// TwinCAT 3 PLC project PLCLibrary
// Title: LPLC
// Company: LPLC
// Author: Arya Farzin
// ProjectVersion: 2.2.0
// Description: LPLC - standardized TwinCAT 3 device, motion and machine function blocks (companion PLC library to lhmi). MIT License.
// ProgramVersion: 3.1.4026.17
// libraries:
//   Tc2_MC2, * (Beckhoff Automation GmbH)
//   Tc2_MC2_Camming, * (Beckhoff Automation GmbH)
//   Tc2_ModbusSrv, * (Beckhoff Automation GmbH)
//   Tc2_Standard, * (Beckhoff Automation GmbH)
//   Tc2_SUPS, * (Beckhoff Automation GmbH)
//   Tc2_System, * (Beckhoff Automation GmbH)
//   Tc2_Utilities, * (Beckhoff Automation GmbH)
//   Tc3_EventLogger, * (Beckhoff Automation GmbH)
//   Tc3_IotBase, * (Beckhoff Automation GmbH)
//   Tc3_JsonXml, * (Beckhoff Automation GmbH)
// project tree:
//   DUTs/Abstract/abs_fb_Device/ ST_Device_HMI_Interface.TcDUT
//   DUTs/Abstract/abs_fb_stateDevice/ ST_StateDevice_HMI_Commands.TcDUT, ST_StateDevice_HMI_Interface.TcDUT, ST_StateDevice_HMI_Status.TcDUT
//   DUTs/Abstract/abs_fb_MachineFlow/ ST_MachineFlow_HMI_Status.TcDUT, ST_MachineFlow_Step.TcDUT, ST_MachineFlow_Transition.TcDUT
//   DUTs/Devices/fb_Dev_StackLight3SegHV_BannerTL50Pro/ EN_Banner_TL503Pro_Animation.TcDUT, EN_Banner_TL503Pro_Colors.TcDUT, ST_Banner_TL503Pro.TcDUT, ST_Banner_TL503Pro_Raw.TcDUT
//   DUTs/Comm/fb_Modbus_Driver/ E_DriverState.TcDUT, E_MBArea.TcDUT, E_MBDataType.TcDUT, E_SignalQuality.TcDUT, E_WordOrder.TcDUT, ST_BitRegisterRmw.TcDUT, ST_MBDeviceStatus.TcDUT, ST_MBReadResult.TcDUT, ST_MBSignalConfig.TcDUT, ST_MBWriteData.TcDUT, ST_ParsedSignal.TcDUT, ST_ReadBlock.TcDUT, ST_WriteBlock.TcDUT
//   DUTs/Comm/fb_MQTT_Connector/ E_MQTT_Direction.TcDUT, E_MQTT_PublishMode.TcDUT, E_MQTT_SignalType.TcDUT, ST_MQTT_Signal.TcDUT
//   DUTs/Devices/fb_Dev_AnalogSensor/ ST_AnalogSensor_Diag.TcDUT, ST_AnalogSensor_HMI_Interface.TcDUT
//   DUTs/Devices/fb_Dev_IsolationMonitor/ ST_IsoMon_DeviceSignals.TcDUT, ST_IsoMon_HMI_Interface.TcDUT, ST_IsoMon_MBIF.TcDUT
//   DUTs/Devices/fb_Dev_PSU_ITECH/ ST_ITECH_DCMeter.TcDUT, ST_ITECH_DCSource.TcDUT, ST_ITECH_DeviceSignals.TcDUT, ST_ITECH_HMI_DeviceSignals.TcDUT, ST_ITECH_Protection.TcDUT, ST_ITECH_QuestionRegister.TcDUT, ST_ITECH_SetConfigs.TcDUT, ST_ITECH_SoftwareFaults.TcDUT, ST_ITECH_SystemStatus.TcDUT
//   DUTs/Devices/fb_Dev_Pump_ABBACS580/ ST_Pump_ABBACS580_HMI_Interface.TcDUT
//   DUTs/Devices/fb_Dev_Pump_SPAL/ EN_Pump_SPAL_Operating_Status.TcDUT, EN_Pump_SPAL_PumpError.TcDUT, EN_Pump_SPAL_ServiceIndicator.TcDUT, ST_Pump_SPAL_CAN_Inputs.TcDUT, ST_Pump_SPAL_CAN_Outputs.TcDUT, ST_Pump_SPAL_HMI_Interface.TcDUT
//   DUTs/Devices/fb_Dev_Actuator/ ST_Actuator_HMI_Interface.TcDUT
//   DUTs/Devices/fb_Dev_VFD_ABBACS580/ ST_VFD_ABBACS580_HMI_Interface.TcDUT, ST_VFD_ABBACS580_Telemetry.TcDUT
//   DUTs/Devices/fb_Dev_VFD_DuraPulse/ ST_VFD_DuraPulse_HMI_Interface.TcDUT, ST_VFD_DuraPulse_Telemetry.TcDUT
//   DUTs/fb_Axis/ E_Axis_BufferMode.TcDUT, E_Axis_JogSource.TcDUT, E_Axis_Mode.TcDUT, E_Axis_UnitType.TcDUT, ST_Axis_HMI_Commands.TcDUT, ST_Axis_HMI_Config.TcDUT, ST_Axis_HMI_Interface.TcDUT, ST_Axis_HMI_Status.TcDUT, ST_Axis_MoveDefinition.TcDUT
//   DUTs/Camming/fb_CamCoupler/ E_CamCoupler_State.TcDUT, ST_CamCoupler_HMI_Commands.TcDUT, ST_CamCoupler_HMI_Config.TcDUT, ST_CamCoupler_HMI_Interface.TcDUT, ST_CamCoupler_HMI_Status.TcDUT
//   DUTs/Camming/fb_CamTeach/ E_CamTeach_Interp.TcDUT, E_CamTeach_State.TcDUT, ST_CamTeach_HMI_Commands.TcDUT, ST_CamTeach_HMI_Config.TcDUT, ST_CamTeach_HMI_Interface.TcDUT, ST_CamTeach_HMI_Status.TcDUT, ST_CamTeach_Point.TcDUT
//   DUTs/Devices/fb_Dev_StripLight_BannerWLS15Pro/ E_BannerWLS15Pro_Animation.TcDUT, E_BannerWLS15Pro_Color.TcDUT, E_BannerWLS15Pro_Direction.TcDUT, E_BannerWLS15Pro_Intensity.TcDUT, E_BannerWLS15Pro_PulsePattern.TcDUT, E_BannerWLS15Pro_ScrollBounceStyle.TcDUT, E_BannerWLS15Pro_Speed.TcDUT, ST_Banner_WLS15PXRGB0220DSKQP_RunMode_Outputs.TcDUT
//   DUTs/Devices/fb_Dev_XPendant/ ST_XPendant_Axis.TcDUT, ST_XPendant_HMI_Interface.TcDUT, ST_XPendant_HMI_Status.TcDUT, ST_XPendant_In.TcDUT
//   DUTs/Common/ ST_Bits.TcDUT, U_ByteToLReal.TcDUT, U_UINT16.TcDUT, U_USINT.TcDUT
//   DUTs/Devices/fb_Dev_ControlValve_Modulating/ ST_ControlValve_Modulating_HMI_Interface.TcDUT
//   DUTs/fb_IO_EL6751_Bus_Status/ ST_EL6751_Bus_State.TcDUT, ST_EL6751_Bus_State_Parsed.TcDUT
//   DUTs/fb_Interlock/ ST_Interlock.TcDUT, ST_Interlock_HMI_Interface.TcDUT
//   DUTs/fb_Permissive/ ST_Permissive.TcDUT, ST_Permissive_HMI_Interface.TcDUT
//   DUTs/fb_Machine/ ST_Machine_HMI_Interface.TcDUT
//   DUTs/Comm/ ST_Modbus_Commands.TcDUT, ST_Modbus_Device_Config.TcDUT
//   POUs/FBs/Abstract/ abs_fb_Device.TcPOU, abs_fb_MachineFlow.TcPOU, abs_fb_stateDevice.TcPOU
//   POUs/FBs/Comm/ fb_Modbus_Driver.TcPOU, fb_MQTT_Connector.TcPOU
//   POUs/FBs/ fb_WriteDataToFile.TcPOU, fb_Axis.TcPOU, fb_FaultMonitor.TcPOU, fb_HmiEventLog.TcPOU, fb_Interlock.TcPOU, fb_Permissive.TcPOU, fb_IO_EL6751_Bus_Status.TcPOU, fb_Machine.TcPOU, fb_PID_Clamping.TcPOU, fb_RampGenerator.TcPOU, fb_SampleBuffer.TcPOU, fb_TimeAverage.TcPOU
//   POUs/FBs/Devices/ fb_Dev_Actuator.TcPOU, fb_Dev_XPendant.TcPOU, fb_Dev_AnalogSensor.TcPOU, fb_Dev_AnalogSensor_Accelerometer.TcPOU, fb_Dev_AnalogSensor_CurrentTransducer.TcPOU, fb_Dev_AnalogSensor_ELM_10x.TcPOU, fb_Dev_AnalogSensor_ELM_10x_CurrentTransducer.TcPOU, fb_Dev_ControlValve_Modulating_INT.TcPOU, fb_Dev_Pump_ABBACS580.TcPOU, fb_Dev_VFD_ABBACS580.TcPOU, fb_Dev_VFD_DuraPulse.TcPOU, fb_Dev_WebRelay.TcPOU, fb_Dev_ControlValve_Modulating.TcPOU, fb_Dev_ControlValve_Modulating_REAL.TcPOU, fb_Dev_IsolationMonitor.TcPOU, fb_Dev_Machine.TcPOU, fb_Dev_PSU_ITECH.TcPOU, fb_Dev_Pump_SPAL.TcPOU, fb_Dev_StackLight3SegHV_BannerTL50Pro.TcPOU, fb_Dev_StripLight_BannerWLS15Pro.TcPOU
//   POUs/FBs/Camming/ fb_CamCoupler.TcPOU, fb_CamTeach.TcPOU, fb_CamTeachFile.TcPOU
//   POUs/FC/ F_AddToArray_String.TcPOU, F_AnalogToEngUnit.TcPOU, F_RemoveFromArray_String.TcPOU
//   GVLs/ GVL_Cam.TcGVL
//   Version/ Global_Version.TcGVL

// ---- DUTs/Abstract/abs_fb_Device/ST_Device_HMI_Interface.TcDUT
TYPE ST_Device_HMI_Interface :
STRUCT
	enabled				: BOOL;
	deviceName			: STRING;
	interlock			: ST_Interlock_HMI_Interface;
	stsInAuto			: BOOL;
	stsFaulted			: BOOL;
	stsFaultDescription	: STRING;
END_STRUCT
END_TYPE

// ---- DUTs/Abstract/abs_fb_stateDevice/ST_StateDevice_HMI_Commands.TcDUT
TYPE ST_StateDevice_HMI_Commands :
STRUCT
	ocmdRun				: BOOL;
	ocmdReset			: BOOL;
	ocmdAbort			: BOOL;
	ocmdRetry			: BOOL;
END_STRUCT
END_TYPE

// ---- DUTs/Abstract/abs_fb_stateDevice/ST_StateDevice_HMI_Interface.TcDUT
TYPE ST_StateDevice_HMI_Interface :
STRUCT
	Status		: ST_StateDevice_HMI_Status;
	Commands 	: ST_StateDevice_HMI_Commands;
	Interlock  	: ST_Interlock_HMI_Interface;
	// Conditions that must be met for this device to ENTER Running (cmdSetStartPermissive). Purely
	// ADDITIVE — a device that never wires a slot publishes an all-satisfied permissive, so nothing
	// that read this struct before needs to change.
	startPermissive	: ST_Permissive_HMI_Interface;

END_STRUCT
END_TYPE

// ---- DUTs/Abstract/abs_fb_stateDevice/ST_StateDevice_HMI_Status.TcDUT
TYPE ST_StateDevice_HMI_Status :
STRUCT
	cfgDeviceName		: STRING;
	stsAuto				: BOOL;
	stsIdle				: BOOL;
	stsDone				: BOOL;
	stsRunning 			: BOOL;
	stsFaulted			: BOOL;
	stsAborting			: BOOL;
	stsAborted			: BOOL;
	stsFaultDescription	: STRING;
	stsState			: STRING;
	stsStepDescription	: STRING;
	stsStepNumber		: INT;
	stsRetryAllowed		: BOOL;
END_STRUCT
END_TYPE

// ---- DUTs/Abstract/abs_fb_MachineFlow/ST_MachineFlow_HMI_Status.TcDUT
// HMI status published by abs_fb_MachineFlow (member HMIflow / getFlowHMIdata()).
// Complements the inherited ST_StateDevice_HMI_Interface (state/step/commands):
// this struct carries what a flow-chart renderer needs. The token masks are two
// UDINT halves (not one LWORD) so a JSON/JS transport never exceeds 2^53.
// stsFlowDef is STATIC after startup - read it once, on demand, not cyclically.
TYPE ST_MachineFlow_HMI_Status :
STRUCT
    stsActiveLo    : UDINT;   // token mask, steps 1..32 (bit = step id - 1)
    stsActiveHi    : UDINT;   // token mask, steps 33..64 (bit = step id - 33)
    stsDoneLo      : UDINT;   // done-and-waiting mask (subset of active), steps 1..32
    stsDoneHi      : UDINT;   // done-and-waiting mask, steps 33..64
    stsPermissiveLo : UDINT;   // permissive mask, transitions 1..32 (bit set = permissive MET)
    stsPermissiveHi : UDINT;   // permissive mask, transitions 33..64
    // HISTORY for this run, cleared on run/reset. Without these an HMI cannot tell a step that
    // COMPLETED from one that never ran - both simply have no token - nor which transitions fired
    // beyond the most recent one. The flow chart needs that distinction to colour progress:
    // active / completed / never-reached are three different things to an operator.
    stsVisitedLo   : UDINT;   // steps whose token was consumed by a firing transition, 1..32
    stsVisitedHi   : UDINT;   // ditto, steps 33..64
    stsFiredLo     : UDINT;   // transitions that have FIRED this run, 1..32 (stsLastFired is only the newest)
    stsFiredHi     : UDINT;   // ditto, transitions 33..64
    // Step id that owns the active fault, 0 = none. Covers BOTH routes: a step body calling
    // setFault() on the inherited state device (the step is stateful, so the fault belongs to it),
    // and a step timeout. First claim wins, so a later step in the same scan cannot steal it.
    stsFaultedStep : INT;
    stsFireCount   : INT;     // transition firings this run (mirrors the base stsStepNumber)
    stsLastFired   : INT;     // last transition id fired; 0 = none
    stsStepCount   : INT;
    stsTransCount  : INT;
    stsActiveNames : STRING(255);   // ' + '-joined names of the active steps
    stsFlowDef     : STRING(4095);   // the graph as JSON: {"v":1,"steps":[{"i","n","d","init"}],"trans":[{"id","n","s":[],"t":[]}]}
END_STRUCT
END_TYPE

// ---- DUTs/Abstract/abs_fb_MachineFlow/ST_MachineFlow_Step.TcDUT
// One step of an abs_fb_MachineFlow sequence. Declared via addStep(); the
// runtime members are ENGINE-OWNED (step bodies use stepDone()/stepElapsed(),
// never these members directly).
TYPE ST_MachineFlow_Step :
STRUCT
    name        : STRING(63);    // shown on the HMI; no double quotes (embedded in the def JSON)
    description : STRING(125);   // WHAT the step does - shown in the HMI's step popup; no double quotes
    timeout     : TIME;          // T#0S = none; engine faults (retryable) when elapsed exceeds it
    active      : BOOL;         // token present
    done        : BOOL;         // step body reported complete; cleared when a transition consumes the token
    entered     : BOOL;         // step body has run at least one scan since activation
    kickTimer   : BOOL;         // one-scan request to restart the step's elapsed clock
    hasOutgoing : BOOL;         // derived from the transitions; done + terminal => sequence Done
    visited    : BOOL;   // completed at least once this run (token consumed by a firing transition)
END_STRUCT
END_TYPE

// ---- DUTs/Abstract/abs_fb_MachineFlow/ST_MachineFlow_Transition.TcDUT
// One transition of an abs_fb_MachineFlow sequence - the ONLY relationship
// object between steps. Fires when ALL source steps are active AND done AND
// the permissive is TRUE; firing consumes the source tokens and activates all
// targets. 1->N = AND-divergence, N->1 = AND-convergence, two transitions from
// one step with opposing permissives = OR-choice, a backward target = a loop.
TYPE ST_MachineFlow_Transition :
STRUCT
    name       : STRING(63);   // the CONDITION text shown on the HMI (e.g. 'cycles < 3'); no double quotes
    sources    : ARRAY[1..4] OF INT;   // step ids; 0 = unused slot
    targets    : ARRAY[1..4] OF INT;   // step ids; 0 = unused slot
    // The gate, and the ONLY thing the engine knows about it. Set with setPermissive(); sticky, and
    // reset to TRUE on reset. Where the gate is really an fb_Permissive, the machine ANDs it in at
    // the call site — setPermissive(t, PermUnload.stsPermissiveOK) — exactly as it reports a step
    // with stepDone(id). An earlier revision carried a POINTER TO fb_Permissive here instead, so the
    // engine dereferenced an object it did not own on every scan; removed 2026-07-26, because the
    // boolean already expresses the effective gate, the HMI reads each permissive's conditions
    // straight from that instance, and a stored pointer can go stale where a value cannot.
    permissive : BOOL := TRUE;
    fired      : BOOL;   // has fired at least once this run (reset with the run)
END_STRUCT
END_TYPE

// ---- DUTs/Devices/fb_Dev_StackLight3SegHV_BannerTL50Pro/EN_Banner_TL503Pro_Animation.TcDUT
{attribute 'qualified_only'}
{attribute 'strict'}
{attribute 'to_string'}
TYPE EN_Banner_TL503Pro_Animation :
(
	Off,
	Steady,
	Flash,
	TwoColorFlash,
	FiftyFifty,
	FiftyFiftyRotate,
	Chase,
	IntensitySweep,
	Scroll,
	Bounce,
	ColorSprectrum,
	Demo
);
END_TYPE

// ---- DUTs/Devices/fb_Dev_StackLight3SegHV_BannerTL50Pro/EN_Banner_TL503Pro_Colors.TcDUT
{attribute 'qualified_only'}
{attribute 'strict'}
{attribute 'to_string'}
TYPE EN_Banner_TL503Pro_Colors :
(
	Green,
	Red,
	Orange,
	Amber,
	Yellow,
	LimeGreen,
	SpringGreen,
	Cyan,
	SkyBlue,
	Blue,
	Violet,
	Magenta,
	Rose,
	White,
	Custom1,
	Custom2	
);
END_TYPE

// ---- DUTs/Devices/fb_Dev_StackLight3SegHV_BannerTL50Pro/ST_Banner_TL503Pro.TcDUT
TYPE ST_Banner_TL503Pro:
STRUCT
	Segment1Color1 			: U_USINT;
	Segment1Color1Intensity : U_USINT;
	Segment1AnimationType	: U_USINT;
	Segment1Speed			: U_USINT;
	Segment1PulsePattern	: U_USINT;
	Segment1Color2			: U_USINT;
	Segment1Color2Intensity : U_USINT;
	Segment1RotationDir		: BOOL;
	
	Segment2Color1 			: U_USINT;
	Segment2Color1Intensity : U_USINT;
	Segment2AnimationType	: U_USINT;
	Segment2Speed			: U_USINT;
	Segment2PulsePattern	: U_USINT;
	Segment2Color2			: U_USINT;
	Segment2Color2Intensity : U_USINT;
	Segment2RotationDir		: BOOL;
	
	Segment3Color1 			: U_USINT;
	Segment3Color1Intensity : U_USINT;
	Segment3AnimationType	: U_USINT;
	Segment3Speed			: U_USINT;
	Segment3PulsePattern	: U_USINT;
	Segment3Color2			: U_USINT;
	Segment3Color2Intensity : U_USINT;
	Segment3RotationDir	: BOOL;
	
END_STRUCT
END_TYPE

// ---- DUTs/Devices/fb_Dev_StackLight3SegHV_BannerTL50Pro/ST_Banner_TL503Pro_Raw.TcDUT
TYPE ST_Banner_TL503Pro_Raw :
STRUCT
	PDOs	:	Array[20..30] of USINT;
END_STRUCT
END_TYPE

// ---- DUTs/Comm/fb_Modbus_Driver/E_DriverState.TcDUT
{attribute 'qualified_only'}
{attribute 'strict'}
TYPE E_DriverState :
(
    Init                := 0,
    ParseConfig         := 1,
    OptimizeBlocks      := 2,

    Connecting          := 5,
    ConnectWait         := 6,
    Ready               := 10,

    ReadStart           := 20,
    ReadSend            := 21,
    ReadWait            := 22,
    ReadProcess         := 23,
    ReadDelay           := 24,
    ReadComplete        := 29,

    WriteStart          := 30,
    WriteSend           := 31,
    WriteWait           := 32,
    WriteDelay          := 33,
    WriteComplete       := 39,

    RmwReadSend         := 40,
    RmwReadWait         := 41,
    RmwModify           := 42,
    RmwWriteSend        := 43,
    RmwWriteWait        := 44,
    RmwDelay            := 45,

    Disconnecting       := 80,
    DisconnectWait      := 81,
    ReconnectWait       := 85,

    Error               := 90,
    Faulted             := 99
) UINT;
END_TYPE

// ---- DUTs/Comm/fb_Modbus_Driver/E_MBArea.TcDUT
{attribute 'qualified_only'}
{attribute 'strict'}
TYPE E_MBArea :
(
    Coils               := 0,
    DiscreteInputs      := 1,
    InputRegisters      := 3,
    HoldingRegisters    := 4
) UINT;
END_TYPE

// ---- DUTs/Comm/fb_Modbus_Driver/E_MBDataType.TcDUT
{attribute 'qualified_only'}
{attribute 'strict'}
{attribute 'to_string'}
TYPE E_MBDataType :
(
    mbNone      := 0,
    mbReal32    := 1,
    mbInt32     := 2,
    mbUInt32    := 3,
    mbInt16     := 4,
    mbUInt16    := 5,
    mbWord16    := 6,
    mbBit       := 7
) UINT;
END_TYPE

// ---- DUTs/Comm/fb_Modbus_Driver/E_SignalQuality.TcDUT
{attribute 'qualified_only'}
{attribute 'strict'}
TYPE E_SignalQuality :
(
    Good                := 0,
    BadComm             := 1,
    BadConfig           := 2,
    BadDeviceFault      := 3,
    UncertainStale      := 4,
    UncertainInit       := 5
) UINT;
END_TYPE

// ---- DUTs/Comm/fb_Modbus_Driver/E_WordOrder.TcDUT
{attribute 'qualified_only'}
{attribute 'strict'}
{attribute 'to_string'}
TYPE E_WordOrder :
(
    BigEndian       := 0,
    LittleEndian    := 1
) UINT;
END_TYPE

// ---- DUTs/Comm/fb_Modbus_Driver/ST_BitRegisterRmw.TcDUT
TYPE ST_BitRegisterRmw :
STRUCT
    address             : UINT;
    managedBitMask      : WORD;
    arrSignalIndex      : ARRAY[0..15] OF UINT;
    readValue           : WORD;
    writeValue          : WORD;
END_STRUCT
END_TYPE

// ---- DUTs/Comm/fb_Modbus_Driver/ST_MBDeviceStatus.TcDUT
TYPE ST_MBDeviceStatus :
STRUCT
    connected               : BOOL;
    faulted                 : BOOL;
    readCycleActive         : BOOL;
    writeCycleActive        : BOOL;

    consecutiveFailures     : UINT;
    reconnectAttempts       : UINT;
    totalReadCycles         : UDINT;
    totalWriteCycles        : UDINT;
    totalErrors             : UDINT;

    lastErrorCode           : UDINT;
    timeSinceLastGoodRead   : TIME;
    timeSinceLastGoodWrite  : TIME;

    currentState            : E_DriverState;
    readBlockCount          : UINT;
    writeBlockCount         : UINT;
    bitRegisterCount        : UINT;
END_STRUCT
END_TYPE

// ---- DUTs/Comm/fb_Modbus_Driver/ST_MBReadResult.TcDUT
TYPE ST_MBReadResult :
STRUCT
    valueReal           : REAL;
    valueDint           : DINT;
    valueUdint          : UDINT;
    valueInt            : INT;
    valueUint           : UINT;
    valueWord           : WORD;
    valueBool           : BOOL;

    quality             : E_SignalQuality := E_SignalQuality.UncertainInit;
    updateCount         : UDINT;
END_STRUCT
END_TYPE

// ---- DUTs/Comm/fb_Modbus_Driver/ST_MBSignalConfig.TcDUT
TYPE ST_MBSignalConfig :
STRUCT
    modbusAddr          : UDINT;
    dataType            : E_MBDataType;
    bitIndex            : BYTE := 255;
    tag                 : STRING(32);
END_STRUCT
END_TYPE

// ---- DUTs/Comm/fb_Modbus_Driver/ST_MBWriteData.TcDUT
TYPE ST_MBWriteData :
STRUCT
    valueReal           : REAL;
    valueDint           : DINT;
    valueUdint          : UDINT;
    valueInt            : INT;
    valueUint           : UINT;
    valueWord           : WORD;
    valueBool           : BOOL;

    writeSuccess        : BOOL;
    writeError          : BOOL;
    writeCount          : UDINT;
END_STRUCT
END_TYPE

// ---- DUTs/Comm/fb_Modbus_Driver/ST_ParsedSignal.TcDUT
TYPE ST_ParsedSignal :
STRUCT
    area                : E_MBArea;
    baseAddress         : UINT;
    bitIndex            : BYTE;
    registerCount       : UINT;
    dataType            : E_MBDataType;
    valid               : BOOL;
    isBitInRegister     : BOOL;
END_STRUCT
END_TYPE

// ---- DUTs/Comm/fb_Modbus_Driver/ST_ReadBlock.TcDUT
TYPE ST_ReadBlock :
STRUCT
    startAddress        : UINT;
    quantity            : UINT;
    area                : E_MBArea;
    functionCode        : BYTE;

    arrSignalIndex      : ARRAY[1..64] OF UINT;
    arrOffsetInBlock    : ARRAY[1..64] OF UINT;
    signalCount         : UINT;

    enabled             : BOOL := TRUE;
END_STRUCT
END_TYPE

// ---- DUTs/Comm/fb_Modbus_Driver/ST_WriteBlock.TcDUT
TYPE ST_WriteBlock :
STRUCT
    startAddress        : UINT;
    quantity            : UINT;
    area                : E_MBArea;
    functionCode        : BYTE;

    arrSignalIndex      : ARRAY[1..64] OF UINT;
    arrOffsetInBlock    : ARRAY[1..64] OF UINT;
    signalCount         : UINT;

    enabled             : BOOL := TRUE;
    containsBitSignals  : BOOL;
END_STRUCT
END_TYPE

// ---- DUTs/Comm/fb_MQTT_Connector/E_MQTT_Direction.TcDUT
// ═══════════════════════════════════════════════════════════════════════
// E_MQTT_Direction - Data flow direction
// ═══════════════════════════════════════════════════════════════════════
{attribute 'qualified_only'}
{attribute 'strict'}
TYPE E_MQTT_Direction :
(
    PUBLISH       := 1,     // PLC → MQTT only
    SUBSCRIBE     := 2,     // MQTT → PLC only  
    BIDIRECTIONAL := 3      // Both directions
);
END_TYPE

// ---- DUTs/Comm/fb_MQTT_Connector/E_MQTT_PublishMode.TcDUT
// ═══════════════════════════════════════════════════════════════════════
// E_MQTT_PublishMode - When to publish
// ═══════════════════════════════════════════════════════════════════════
{attribute 'qualified_only'}
{attribute 'strict'}
TYPE E_MQTT_PublishMode :
(
    DISABLED            := 0,   // Don't publish (subscribe-only signal)
    CHANGE_OF_STATE     := 1,   // Publish only when value changes
    PERIODIC            := 2,   // Publish at fixed interval (also publishes on change)
    TRANSACTION_GROUP_1 := 3,   // Grouped JSON publish (default 100ms period)
    TRANSACTION_GROUP_2 := 4,   // Grouped JSON publish (default 1s period)
    TRANSACTION_GROUP_3 := 5    // Grouped JSON publish (default 5s period)
);
END_TYPE

// ---- DUTs/Comm/fb_MQTT_Connector/E_MQTT_SignalType.TcDUT
// ═══════════════════════════════════════════════════════════════════════
// E_MQTT_SignalType - Supported data types for MQTT signals
// ═══════════════════════════════════════════════════════════════════════
{attribute 'qualified_only'}
{attribute 'strict'}
TYPE E_MQTT_SignalType :
(
    NONE        := 0,
    TYPE_BOOL   := 1,
    TYPE_BYTE   := 2,
    TYPE_INT    := 3,
    TYPE_DINT   := 4,
    TYPE_REAL   := 5,
    TYPE_LREAL  := 6,
    TYPE_STRING := 7,
    TYPE_TIME   := 8
);
END_TYPE

// ---- DUTs/Comm/fb_MQTT_Connector/ST_MQTT_Signal.TcDUT
// ═══════════════════════════════════════════════════════════════════════
// ST_MQTT_Signal - Internal signal descriptor
// ═══════════════════════════════════════════════════════════════════════
TYPE ST_MQTT_Signal :
STRUCT
    // Configuration (set by user during registration)
    sSubTopic           : STRING(80);           // Topic suffix, e.g. 'PIT1/stsEngValue'
    pValue              : PVOID;                // Pointer to the PLC variable
    eType               : E_MQTT_SignalType;    // Data type for serialization
    ePublishMode        : E_MQTT_PublishMode;   // CoS or Periodic
    eDirection          : E_MQTT_Direction;     // Pub / Sub / Both
    tPublishInterval    : TIME;                 // Interval for PERIODIC mode
    sJsonKey            : STRING(255);          // JSON key to extract (empty = raw payload mode)
    sJsonParentKey      : STRING(80);           // Optional parent object key (e.g. 'signals')
    
    // Internal state (managed by FB)
    sLastPublished      : STRING(255);          // Last published value (for CoS detection)
    tLastPublishTime    : TIME;                 // Timestamp of last publish
    bRegistered         : BOOL;                 // TRUE if this slot is in use
    nConsecFails        : UINT;                 // Consecutive failures for this signal
END_STRUCT
END_TYPE

// ---- DUTs/Devices/fb_Dev_AnalogSensor/ST_AnalogSensor_Diag.TcDUT
TYPE ST_AnalogSensor_Diag :
STRUCT
	NoOfSamples : USINT;
	error		: BIT;
	underrange	: BIT;
	overrange	: BIT;
	diag		: BIT;
	limit1		: BIT;
	limit2		: BIT;

END_STRUCT
END_TYPE

// ---- DUTs/Devices/fb_Dev_AnalogSensor/ST_AnalogSensor_HMI_Interface.TcDUT
TYPE ST_AnalogSensor_HMI_Interface :
STRUCT
	HMIbaseDevice		: ST_Device_HMI_Interface;
	stsSensorRawSignal	: LREAL;
	stsEngValue			: LREAL;
	cfgAlarmEnable		: BOOL;
	cfgAlarmL			: LREAL;
	cfgAlarmLL			: LREAL;
	cfgAlarmH			: LREAL;
	cfgAlarmHH			: LREAL;
	cfgEngUnit			: STRING;
	cfgCalOffset		: LREAL;
	cfgCalGain			: LREAL;
END_STRUCT
END_TYPE

// ---- DUTs/Devices/fb_Dev_IsolationMonitor/ST_IsoMon_DeviceSignals.TcDUT
TYPE ST_IsoMon_DeviceSignals :
STRUCT
	insulationResistance_kOhm : REAL;
	minInsulationValue	 	: REAL;
	voltageDCPlusToMinus 	: REAL;
	voltageDCPlusToPE	 	: REAL;
	voltageDCMinusToPE	 	: REAL;
	couplingToSystem	 	: REAL;
	couplingtoEarth		 	: REAL;
	deviceError			 	: REAL;
	deviceInactive			: REAL;
	dcOffset				: REAL;
	measurementQuality		: REAL;
END_STRUCT
END_TYPE

// ---- DUTs/Devices/fb_Dev_IsolationMonitor/ST_IsoMon_HMI_Interface.TcDUT
TYPE ST_IsoMon_HMI_Interface :
STRUCT
	HMIbaseDevice		: ST_Device_HMI_Interface; 
	ocmdTripReset		: BOOL;
	ocmdTest			: BOOL;
	stsDeviceAlarm		: BOOL;
	stsDeviceWarning	: BOOL;
END_STRUCT
END_TYPE

// ---- DUTs/Devices/fb_Dev_IsolationMonitor/ST_IsoMon_MBIF.TcDUT
TYPE ST_IsoMon_MBIF :
STRUCT
    insulationResistance      : U_ByteToLReal;   // 0x2000: Insulation resistance in Ω
    minInsulationValue        : U_ByteToLReal;   // 0x2002: Minimum insulation resistance in Ω
    systemLeakageCapacitance  : U_ByteToLReal;   // 0x2004: System leakage capacitance in F
    voltageL1L2               : U_ByteToLReal;   // 0x2006: Voltage from phase L1 to phase L2 in V
    voltageL1L3               : U_ByteToLReal;   // 0x2008: Voltage from phase L1 to phase L3 in V
    voltageL2L3               : U_ByteToLReal;   // 0x200A: Voltage from phase L2 to phase L3 in V
    voltageL1PE               : U_ByteToLReal;   // 0x200C: Voltage from phase L1 to earth PE in V
    voltageL2PE               : U_ByteToLReal;   // 0x200E: Voltage from phase L2 to earth PE in V
    voltageL3PE               : U_ByteToLReal;   // 0x2010: Voltage from phase L3 to earth PE in V
    systemFrequency           : U_ByteToLReal;   // 0x2012: System frequency in Hz
    couplingToSystem          : U_ByteToLReal;   // 0x2014: Coupling to system (0 = O.K., 101 = fault)
    couplingToEarth           : U_ByteToLReal;   // 0x2016: Coupling to earth (0 = O.K., 102 = fault)
    deviceError               : U_ByteToLReal;   // 0x2018: Device error number (example: 750 -> 750 communication CAN)
    deviceInactive            : U_ByteToLReal;   // 0x201A: Device inactive (0 = active, 1 = inactive)
    dcOffset                  : U_ByteToLReal;   // 0x201C: DC offset in the system (0..100%) in %
    measurementQuality        : U_ByteToLReal;   // 0x201E: Measured value quality (0% = bad, 100% = good) in %
    symmetricalAlarm          : U_ByteToLReal;   // 0x2020: Symmetrical alarm (see 0x1121)
    dcMinusAlarm              : U_ByteToLReal;   // 0x2022: DC- alarm (see 0x1121)
    dcPlusAlarm               : U_ByteToLReal;   // 0x2024: DC+ alarm (see 0x1121)
    durationMeasuringPulse    : U_ByteToLReal;   // 0x2026: Duration of the measuring pulse (0% = short, 100% = long) in %
    voltageDCPE               : U_ByteToLReal;   // 0x2028: DC offset voltage to earth in V
END_STRUCT
END_TYPE

// ---- DUTs/Devices/fb_Dev_PSU_ITECH/ST_ITECH_DCMeter.TcDUT
TYPE ST_ITECH_DCMeter :
STRUCT
	DCVrms      : REAL;   // DC-METER: v_rms (float)
    DCIrms      : REAL;   // DC-METER: i_rms (float)
    DCPrms      : REAL;   // DC-METER: p_rms (float)
    DCOperReg   : UDINT;  // DC-METER: oper_reg (uint32)
    DCStateReg  : UDINT;  // DC-METER: state_reg (uint32)
    DCQuesReg   : UDINT;  // DC-METER: ques_reg (uint32)
    DCSenseVolt : REAL;   // DC-METER: sense_volt (float)
END_STRUCT
END_TYPE

// ---- DUTs/Devices/fb_Dev_PSU_ITECH/ST_ITECH_DCSource.TcDUT
TYPE ST_ITECH_DCSource :
STRUCT
	DCMode			  : UDINT;
	DCVoltSP		  : REAL;
	DCVoltRise		  : REAL;
	DCVoltFall		  : REAL;
	DCCurrentSP		  : REAL;
	DCCurrentRise	  : REAL;
	DCCurrentFall	  : REAL;
	DCVoltHigh        : REAL;   // dc_v_high (float)
    DCVoltLow         : REAL;   // dc_v_low (float)
    DCCurrentHigh     : REAL;   // dc_i_high (float)
    DCCurrentLow      : REAL;   // dc_i_low (float)
    DCCC_SpeedState   : UDINT;  // cc_speed_state (uint32)
    DCCV_SpeedState   : UDINT;  // cv_speed_state (uint32)
    DCPowerHigh       : REAL;   // power_high (float)
    DCPowerLow        : REAL;   // power_low (float)
    DCSlewMode        : UDINT;  // Slew mode (uint32)
    DCOnlyLoad        : UDINT;  // Only Load (uint32)
    DCBatterySim      : UDINT;  // Battery Simulation (uint32)
END_STRUCT
END_TYPE

// ---- DUTs/Devices/fb_Dev_PSU_ITECH/ST_ITECH_DeviceSignals.TcDUT
TYPE ST_ITECH_DeviceSignals :
STRUCT
	DCMeter		:ST_ITECH_DCMeter;
	DCSource	:ST_ITECH_DCSource;
	Protection	:ST_ITECH_Protection;
	System		:ST_ITECH_SystemStatus;
END_STRUCT
END_TYPE

// ---- DUTs/Devices/fb_Dev_PSU_ITECH/ST_ITECH_HMI_DeviceSignals.TcDUT
TYPE ST_ITECH_HMI_DeviceSignals :
STRUCT
	deviceSignals_read	: ST_ITECH_DeviceSignals;
	deviceSignals_write	: ST_ITECH_DeviceSignals;
END_STRUCT
END_TYPE

// ---- DUTs/Devices/fb_Dev_PSU_ITECH/ST_ITECH_Protection.TcDUT
TYPE ST_ITECH_Protection :
STRUCT

    OVPState     : UDINT;  // OVP_state (uint32)
    OVPLevel     : REAL;   // OVP_level (float)
    OVPDelay     : REAL;   // OVP_delay (float)
    OCPState     : UDINT;  // OCP_state (uint32)
 	OCPLevel     : REAL;   // OCP_level (float)
    OCPDelay     : REAL;   // OCP_delay (float)
    OPPState     : UDINT;  // OPP_state (uint32)
    OPPLevel     : REAL;   // OPP_level (float)
    OPPDelay     : REAL;   // OPP_delay (float)
    UCPState     : UDINT;  // UCP_state (uint32)
    UCPLevel     : REAL;   // UCP_level (float)
    UCPDelay     : REAL;   // UCP_delay (float)
    UCPWarmup    : REAL;   // UCP_warmup (float)
    UVPState     : UDINT;  // UVP_state (uint32)
    UVPLevel     : REAL;   // UVP_level (float)
    UVPDelay     : REAL;   // UVP_delay (float)
    UVPWarmup    : REAL;   // UVP_warmup (float)
END_STRUCT
END_TYPE

// ---- DUTs/Devices/fb_Dev_PSU_ITECH/ST_ITECH_QuestionRegister.TcDUT
TYPE ST_ITECH_QuestionRegister :
STRUCT
	overVoltageProtection : BOOL;
	overCurrentProtection : BOOL;
	overPowerProtection	  : BOOL;
	underVoltageProtection: BOOL;
	overTempProtection	  : BOOL;
	underCurrentProtection: BOOL;
	senseFault			  : BOOL;
	currentSharingFault   : BOOL;
	reserved			  : BOOL;
	externalInhibit		  : BOOL;
	faultProtection		  : BOOL;
	loopOscFailure		  : BOOL;
	outputNotRegulated    : BOOL;
END_STRUCT
END_TYPE

// ---- DUTs/Devices/fb_Dev_PSU_ITECH/ST_ITECH_SetConfigs.TcDUT
TYPE ST_ITECH_SetConfigs :
STRUCT
	dcSource	: ST_ITECH_DCSource;
	protection	: ST_ITECH_Protection;
END_STRUCT
END_TYPE

// ---- DUTs/Devices/fb_Dev_PSU_ITECH/ST_ITECH_SoftwareFaults.TcDUT
TYPE ST_ITECH_SoftwareFaults :
STRUCT
	overVoltageProtection 				: BOOL;
	positiveOverCurrentProtection 		: BOOL;
	negativeOverCurrentProtection 		: BOOL;
	positiveOverPowerProtection	 		: BOOL;
	negativeOverPowerProtection  		: BOOL;
	underCurrentProtection		 		: BOOL;
	underVoltageProtection				: BOOL;
	overTemperatureProtection			: BOOL;
	senseAbnormal						: BOOL;
	senseReverseProtection 				: BOOL;
	outputReverseProtection 			: BOOL;
	multiMasterUnitsAbnormal			: BOOL;
	opticalFiberUnlocked_multiMaster	: BOOL;
	opticalFiberUnlocked_singleMaster	: BOOL;
	moduleCheckingFailure				: BOOL;
	unevenCurrentProtection				: BOOL;
	hardwareProtection					: BOOL;
	masterUnitPowerFailureProtection 	: BOOL;
	inhibit_latchmode					: BOOL;
	inhibit_livingMode					: BOOL;
	capacitorOverCurrentprotection		: BOOL;
	slaveUnitPowerFailureProtection		: BOOL;
END_STRUCT
END_TYPE

// ---- DUTs/Devices/fb_Dev_PSU_ITECH/ST_ITECH_SystemStatus.TcDUT
TYPE ST_ITECH_SystemStatus :
STRUCT
	ON_OFF				: UDINT;
	SenseVolt			: REAL;
	Heartbeat			: UDINT;
	Timer_ON_OFF		: UDINT;
	RemoteSenseStatus	: UDINT;
	RemoteSenseLevel	: REAL;
	OutputRZero			: UDINT;
	MeasureCycle		: UDINT;
END_STRUCT
END_TYPE

// ---- DUTs/Devices/fb_Dev_Pump_ABBACS580/ST_Pump_ABBACS580_HMI_Interface.TcDUT
TYPE ST_Pump_ABBACS580_HMI_Interface :
STRUCT
	HMIbaseDevice			: ST_Device_HMI_Interface;
	stsInterlocks			: ST_Interlock_HMI_Interface;

	// Operator commands — pump HMI is the sole command surface when this FB wraps a VFD.
	// (The inner VFD is forced to auto, so VFD.HMI.ocmd* fields are inert.)
	ocmdReset				: BOOL;
	ocmdRun					: BOOL;
	ocmdSetpoint			: LREAL;	// 0..100 percent

	stsOverpressureTripped	: BOOL;
END_STRUCT
END_TYPE

// ---- DUTs/Devices/fb_Dev_Pump_SPAL/EN_Pump_SPAL_Operating_Status.TcDUT
{attribute 'qualified_only'}
{attribute 'strict'}
{attribute 'to_string'}
TYPE EN_Pump_SPAL_Operating_Status :
(
	Normal,
	Derated,
	Not_Operable,
	Not_Available
);
END_TYPE

// ---- DUTs/Devices/fb_Dev_Pump_SPAL/EN_Pump_SPAL_PumpError.TcDUT
{attribute 'qualified_only'}
{attribute 'strict'}
{attribute 'to_string'}
TYPE EN_Pump_SPAL_PumpError :
(
	Normal_Operation,
	Unable_to_start,
	OverV_Protection_Shutdown,
	UnderV_Protection_Shutdown,
	OverT_Protection_Shutdown,
	Speed_Limited_Due_To_Current,
	Speed_Limited_Due_To_Capability,
	Speed_Limited_Due_To_Torque,
	Speed_Limited_Due_To_OverT,
	Reserved1,
	Reserved2,
	Reserved3,
	Reserved4,
	Reserved5,
	Dry_Run	
);
END_TYPE

// ---- DUTs/Devices/fb_Dev_Pump_SPAL/EN_Pump_SPAL_ServiceIndicator.TcDUT
{attribute 'qualified_only'}
{attribute 'strict'}
{attribute 'to_string'}
TYPE EN_Pump_SPAL_ServiceIndicator :
(
   Not_Available,
   Reserved,
   Service_required,
   Service_not_required
);
END_TYPE

// ---- DUTs/Devices/fb_Dev_Pump_SPAL/ST_Pump_SPAL_CAN_Inputs.TcDUT
TYPE ST_Pump_SPAL_CAN_Inputs :
STRUCT
	PumpMotor		: USINT;
	PumpError		: USINT;
	PumpCMDStatus	: USINT;
	PumpSpeed		: LREAL;
	PumpTemperature : LREAL;
	PumpPower		: LREAL;
	PumpServiceIndicator	: USINT;
	PumpOperatorStatus		: USINT;
	
	
	
	
END_STRUCT
END_TYPE

// ---- DUTs/Devices/fb_Dev_Pump_SPAL/ST_Pump_SPAL_CAN_Outputs.TcDUT
TYPE ST_Pump_SPAL_CAN_Outputs :
STRUCT
	MotorStateRequest	: USINT;
	MotorSetpoint		: LREAL;
END_STRUCT
END_TYPE

// ---- DUTs/Devices/fb_Dev_Pump_SPAL/ST_Pump_SPAL_HMI_Interface.TcDUT
TYPE ST_Pump_SPAL_HMI_Interface :
STRUCT
	HMIbaseDevice		: ST_Device_HMI_Interface;
	stsLVOn				: BOOL;
	stsBusStatus		: ST_EL6751_Bus_State_Parsed;
	stsBusOK			: BOOL;
	ocmdReset			: BOOL;
	stsInterlocks		: ST_Interlock_HMI_Interface;
	stsRunPump			: USINT;
	stsSetpoint			: LREAL;

	ocmdRunPump			: USINT;
	ocmdSetpoint		: LREAL;
	stsState			: STRING;
	stsCommandFB		: STRING;
	stsMotorFB			: STRING;
	stsServiceIndicator	: STRING;
	stsError			: STRING;
	stsPower			: LREAL;
	stsTemperature		: LREAL;
	stsSpeed			: LREAL;
		
END_STRUCT
END_TYPE

// ---- DUTs/Devices/fb_Dev_Actuator/ST_Actuator_HMI_Interface.TcDUT
TYPE ST_Actuator_HMI_Interface :
STRUCT
	HMIbaseDevice		: ST_Device_HMI_Interface; 
	stsActuated			: BOOL;
	ocmdActuate			: BOOL;
	ocmdReset			: BOOL;
	setActuate			: BOOL;
END_STRUCT
END_TYPE

// ---- DUTs/Devices/fb_Dev_VFD_ABBACS580/ST_VFD_ABBACS580_HMI_Interface.TcDUT
TYPE ST_VFD_ABBACS580_HMI_Interface :
STRUCT
	HMIbaseDevice		: ST_Device_HMI_Interface;
	stsInterlocks		: ST_Interlock_HMI_Interface;

	// Operator commands
	ocmdReset			: BOOL;
	ocmdRunMode			: USINT;	// 0=stop, 1=fwd, 2=reverse
	ocmdSetpoint		: LREAL;	// percent, -100..+100

	// Command echo
	stsRunMode			: USINT;
	stsSetpoint			: LREAL;

	// Drive state
	stsState			: STRING;
	stsRunning			: BOOL;
	stsAtSetpoint		: BOOL;
	stsRemote			: BOOL;
	stsTripped			: BOOL;
	stsAlarm			: BOOL;

	// Telemetry (engineering units)
	stsActualSpeed		: LREAL;
	stsMotorCurrent		: LREAL;
	stsDCBusVoltage		: LREAL;
	stsOutputFreq		: LREAL;
	stsMotorTorque		: LREAL;
	stsInverterTemp		: LREAL;
	stsFaultCode		: UINT;
	stsFaultText		: STRING;

	// Diagnostics
	stsCWRaw			: WORD;
	stsSWRaw			: WORD;
	stsCommsConnected	: BOOL;
	stsCommsFaulted		: BOOL;
END_STRUCT
END_TYPE

// ---- DUTs/Devices/fb_Dev_VFD_ABBACS580/ST_VFD_ABBACS580_Telemetry.TcDUT
TYPE ST_VFD_ABBACS580_Telemetry :
STRUCT
	actualSpeed		: LREAL;	// percent, signed
	motorCurrent	: LREAL;	// A (raw par 01.07; default whole amps)
	dcBusVoltage	: LREAL;	// VDC (raw 0.1 VDC / 10)
	outputFreq		: LREAL;	// Hz, signed (assumes par 46.02 = 60.0)
	motorTorque		: LREAL;	// %, signed (raw 0.01% / 100)
	inverterTemp	: LREAL;	// % (raw 1%)
	faultCode		: UINT;		// par 04.11 raw
END_STRUCT
END_TYPE

// ---- DUTs/Devices/fb_Dev_VFD_DuraPulse/ST_VFD_DuraPulse_HMI_Interface.TcDUT
TYPE ST_VFD_DuraPulse_HMI_Interface :
STRUCT
	HMIbaseDevice		: ST_Device_HMI_Interface;
	stsInterlocks		: ST_Interlock_HMI_Interface;

	// Operator commands
	ocmdReset			: BOOL;
	ocmdRunMode			: USINT;	// 0=stop, 1=fwd, 2=reverse
	ocmdSetpoint		: LREAL;	// absolute Hz, 0..cfgMaxFreqHz

	// Command echo
	stsRunMode			: USINT;
	stsSetpoint			: LREAL;

	// Drive state
	stsState			: STRING;
	stsRunning			: BOOL;
	stsRemote			: BOOL;
	stsTripped			: BOOL;
	stsAlarm			: BOOL;
	stsDirection		: INT;		// 1=fwd, -1=rev, 0=stopped

	// Telemetry (engineering units)
	stsOutputFreq		: LREAL;	// Hz, signed
	stsMotorRPM			: LREAL;	// rpm, signed
	stsMotorCurrent		: LREAL;	// A
	stsDCBusVoltage		: LREAL;	// VDC
	stsOutputVoltage	: LREAL;	// VAC
	stsMotorTorque		: LREAL;	// %
	stsInverterTemp		: LREAL;	// degC
	stsFaultCode		: USINT;
	stsFaultText		: STRING;
	stsWarningCode		: USINT;
	stsWarningText		: STRING;

	// Diagnostics
	stsCWRaw			: WORD;
	stsSWRaw			: WORD;
	stsCommsConnected	: BOOL;
	stsCommsFaulted		: BOOL;
END_STRUCT
END_TYPE

// ---- DUTs/Devices/fb_Dev_VFD_DuraPulse/ST_VFD_DuraPulse_Telemetry.TcDUT
TYPE ST_VFD_DuraPulse_Telemetry :
STRUCT
	outputFreq		: LREAL;	// Hz, signed (sign reflects direction bits 3-4 of SW)
	motorRPM		: LREAL;	// rpm, signed
	motorCurrent	: LREAL;	// A (raw reg 0x2104 / 100)
	dcBusVoltage	: LREAL;	// VDC (raw reg 0x2105 / 10)
	outputVoltage	: LREAL;	// VAC (raw reg 0x2106 / 10)
	motorTorque		: LREAL;	// % (raw reg 0x210B / 10)
	inverterTemp	: LREAL;	// degC (raw reg 0x220E / 10)
	faultCode		: USINT;	// 0x2100 low byte
	warningCode		: USINT;	// 0x2100 high byte
END_STRUCT
END_TYPE

// ---- DUTs/fb_Axis/E_Axis_BufferMode.TcDUT
TYPE E_Axis_BufferMode :
(
    eAborting     := 0,  // Phase 1 - abort current move, start next immediately
    eBuffered     := 1,  // reserved Phase 2
    eBlendingLow  := 2,  // reserved Phase 2
    eBlendingHigh := 3,  // reserved Phase 2
    eBlendingNext := 4,  // reserved Phase 2
    eBlendingPrev := 5   // reserved Phase 2
) INT;
END_TYPE

// ---- DUTs/fb_Axis/E_Axis_JogSource.TcDUT
// Which input currently owns the jog. HMI jog and the physical teach pendant feed ONE
// MC_Jog through the same gating; this reports/arbitrates which one is in control so the
// two can never command opposite directions. The pendant's dead-man (inpPendantEnable)
// takes ownership while held, locking out the HMI jog buttons.
TYPE E_Axis_JogSource :
(
    eNone    := 0,  // no jog source active
    eHMI     := 1,  // HMI jog buttons
    ePendant := 2   // physical teach pendant (dead-man held)
) INT;
END_TYPE

// ---- DUTs/fb_Axis/E_Axis_Mode.TcDUT
TYPE E_Axis_Mode :
(
    eAbsolute    := 0,  // MC_MoveAbsolute
    eRelative    := 1,  // MC_MoveRelative
    eVelocity    := 2,  // MC_MoveVelocity
    eTorque      := 3,  // MC_TorqueControl
    eHalt        := 4,  // MC_Halt (interruptible)
    eStop        := 5,  // MC_Stop (forced standstill)
    eHome        := 6,  // reserved Phase 2
    eSetPosition := 7,  // reserved Phase 2
    eModulo      := 8,  // absolute target within one modulo period, forced direction (MC_MoveModulo)
    eExternal    := 9   // coordination hook - yields axis to external owner
) INT;
END_TYPE

// ---- DUTs/fb_Axis/E_Axis_UnitType.TcDUT
// Axis kinematic type - drives HMI unit display. NC has no unit metadata, so
// fb_Axis carries this; the actual unit label is configured separately (cfgUnit).
TYPE E_Axis_UnitType :
(
    eLinear := 0,  // translational axis - position e.g. mm, m
    eRotary := 1   // rotational axis  - position e.g. deg, rev
) INT;
END_TYPE

// ---- DUTs/fb_Axis/ST_Axis_HMI_Commands.TcDUT
// HMI → PLC operator commands.
// Move selection is a two-step operation:
//   1. Write ocmdSelectMove (1-20) → stsConfirmPending goes TRUE
//   2. Write ocmdRunMove := TRUE to execute, or ocmdCancelSelect to cancel
TYPE ST_Axis_HMI_Commands :
STRUCT
    ocmdEnable          : BOOL;   // enable axis (power on)
    ocmdDisable         : BOOL;   // disable axis (power off)
    ocmdReset           : BOOL;   // clear faults and release MC_Stop
    ocmdStop            : BOOL;   // forced standstill - locked until reset
    ocmdHome            : BOOL;   // call MC_Home with MC_Direct using HMI.Config.homePosition
    ocmdSelectMove      : INT;    // 1-20: stage a move for confirmation; 0 = no-op
    ocmdRunMove         : BOOL;   // run the staged move (requires a prior ocmdSelectMove)
    ocmdCancelSelect    : BOOL;   // cancel pending selection without executing
    ocmdReloadMoveConfig: BOOL;   // copy persistent live moves -> HMI.Config.moves, discarding un-applied edits
    ocmdApplyMoveConfig : BOOL;   // validate/copy HMI.Config.moves -> persistent live moves when axis is idle
    ocmdJogPositive     : BOOL;   // jog positive direction (level-triggered, hold = continuous)
    ocmdJogNegative     : BOOL;   // jog negative direction (level-triggered, hold = continuous)
    ocmdJogVelocity     : LREAL;  // jog velocity override [unit/s] - 0 = use cfgJogVelocity
    ocmdJogAcceleration : LREAL;  // jog accel override [unit/s²] - 0 = use cfgJogAcceleration
    ocmdVelocityOverride: LREAL;  // velocity override [%] 0-100 - 0 = no change
    // Torque jog: interactive manual torque (dead-man). HOLD ocmdTorqueJog → apply
    // ocmdTorqueJogValue live; release → torque ramps to 0 and the axis stays enabled
    // (free at 0 torque, no MC_Stop). Mutually exclusive with jog/moves/homing.
    ocmdTorqueJog       : BOOL;   // hold = apply torque (level-triggered dead-man)
    ocmdTorqueJogValue  : LREAL;  // live torque setpoint while held [% rated torque]
    ocmdTorqueJogMaxVel : LREAL;  // safety: max |velocity| during torque-jog [unit/s]; 0 = no trip.
                                  // Persistent: retained across restart; FB seeds this field with the
                                  // retained value on the first scan after (re)start (read stsTorqueJogMaxVel).
    // Position jog ("go to position") - a jog subvariant. Write ocmdJogGotoPos with the target
    // (angle or mm), then pulse ocmdJogGoto to run a discrete absolute move at the jog velocity/accel.
    // Mutually exclusive with speed-jog / torque-jog / configured moves / homing.
    ocmdJogGoto         : BOOL;   // run: one-shot, moves to ocmdJogGotoPos (self-cleared by the FB)
    ocmdJogGotoPos      : LREAL;  // [unit] absolute target position (angle or mm)
END_STRUCT
END_TYPE

// ---- DUTs/fb_Axis/ST_Axis_HMI_Config.TcDUT
// HMI-editable axis configuration.
// The move table here is a draft buffer. fb_Axis copies it into the internal
// persistent live move table only when ocmdApplyMoveConfig is accepted.
TYPE ST_Axis_HMI_Config :
STRUCT
    homePosition : LREAL; // position assigned by MC_Home using MC_Direct [unit]
    moves : ARRAY[1..20] OF ST_Axis_MoveDefinition;
END_STRUCT
END_TYPE

// ---- DUTs/fb_Axis/ST_Axis_HMI_Interface.TcDUT
TYPE ST_Axis_HMI_Interface :
STRUCT
    // Inherited base-device HMI values (deviceName, enabled, stsInAuto, stsFaulted,
    // stsFaultDescription, axis-level interlock). Populated from abs_fb_Device.
    HMIbaseDevice : ST_Device_HMI_Interface;
    Status        : ST_Axis_HMI_Status;
    Commands      : ST_Axis_HMI_Commands;
    Config        : ST_Axis_HMI_Config;
END_STRUCT
END_TYPE

// ---- DUTs/fb_Axis/ST_Axis_HMI_Status.TcDUT
TYPE ST_Axis_HMI_Status :
STRUCT
    // Identity, auto mode, fault and axis-level interlock live in HMIbaseDevice
    // (ST_Device_HMI_Interface) - not duplicated here.

    // Axis power state
    stsEnabled          : BOOL;   // MC_Power.Status - drive powered and ready
    stsHomed            : BOOL;   // axis is referenced/calibrated (Axis.Status.Homed)

    // Motion state - curated operator summary (aggregated from AXIS_REF.Status)
    stsStandstill       : BOOL;
    stsMoving           : BOOL;   // DiscreteMotion OR ContinuousMotion
    stsInTargetPos      : BOOL;   // within target window (abs/rel moves)
    stsError            : BOOL;   // NC-level error (separate from PLC fault)
    stsErrorID          : UDINT;  // NC error code

    // Complete AXIS_REF.Status snapshot - every status flag this library version
    // exposes (Disabled, ErrorStop, Stopping, Homing, Homed, DiscreteMotion,
    // ContinuousMotion, SynchronizedMotion, ConstantVelocity, Accelerating,
    // Decelerating, InTargetPosition, ...). Bind this for full/diagnostic status.
    stsAxisStatus       : ST_AxisStatus;

    // Process values
    stsActualPosition   : LREAL;  // [unit]   actual position, accumulated/un-wrapped (Axis.NcToPlc.ActPos)
    // Modulo position - only meaningful when stsIsModulo (the NC axis is configured modulo). The NC
    // computes these regardless, so on a non-modulo axis they are not the value to display.
    stsModuloActPos     : LREAL;  // [unit] actual position wrapped into one modulo period (Axis.NcToPlc.ModuloActPos)
    stsModuloActTurns   : DINT;   // completed modulo turns (Axis.NcToPlc.ModuloActTurns)
    stsActualVelocity   : LREAL;  // [unit/s] actual velocity  (Axis.NcToPlc.ActVelo)
    stsActualTorque     : LREAL;  // [Nm or %] actual torque (Axis.NcToPlc.ActTorque)
    stsSetPosition      : LREAL;  // [unit]   commanded position (Axis.NcToPlc.SetPos)
    stsSetVelocity      : LREAL;  // [unit/s] commanded velocity (Axis.NcToPlc.SetVelo)
    stsSetTorque        : LREAL;  // [% or Nm] commanded torque (FB-tracked; no NC torque setpoint)
    stsFollowingError   : LREAL;  // [unit]   position lag = SetPos - ActPos

    // Homing / direct position assignment
    stsHomeBusy         : BOOL;   // MC_Home.Busy
    stsHomeDone         : BOOL;   // MC_Home.Done
    stsHomeError        : BOOL;   // MC_Home.Error
    stsHomeErrorID      : UDINT;  // MC_Home.ErrorID
    stsHomePosition     : LREAL;  // last/direct home position command [unit]
    stsHomeRetained     : BOOL;   // a taught home is stored and re-applied after restarts (cfgRetainHome)

    // Move status
    stsCurrentMoveIndex : INT;    // 1-20 index of last executed move (0 = none)
    stsCurrentMoveName  : STRING; // moveName of last executed move
    stsMoveBusy         : BOOL;   // MC block is executing
    stsActiveMoveMode   : E_Axis_Mode; // active move mode while stsMoveBusy is TRUE
    stsMoveDone         : BOOL;   // last move completed (position/velocity reached)

    // HMI move selection
    stsSelectedMove     : INT;    // staged move index awaiting confirmation (0 = none)
    stsConfirmPending   : BOOL;   // TRUE: ocmdRunMove required to execute

    // HMI move configuration edit/apply feedback
    stsMoveConfigLoaded     : BOOL;   // TRUE once HMI.Config.moves has been seeded from the live table
    stsMoveConfigApplyError : BOOL;   // last apply/reload command was rejected
    stsMoveConfigErrorText  : STRING; // reason the last apply/reload command was rejected

    // Override
    stsVelocityOverride : LREAL;  // effective velocity override [%] - global value if active, else local
    stsGlobalOverrideActive : BOOL;  // TRUE = axis is following the machine-global override (inpGlobalOverrideEnable)

    // Jog setpoints (currently active - reflects the owning source's velocity/accel)
    stsJogVelocity      : LREAL;  // [unit/s]  active jog velocity
    stsJogAcceleration  : LREAL;  // [unit/s²] active jog acceleration
    stsJogSource        : E_Axis_JogSource;  // which input owns the jog: eNone / eHMI / ePendant
    stsPendantMode      : BOOL;   // teach pendant selected - it owns the jog, HMI jog / torque-jog / go-to locked out
    stsPendantDeadman   : BOOL;   // pendant dead-man held - the pendant can move the axis
    stsJogTorqueLimit   : LREAL;  // [Nm or %] global overtorque trip for position jog (0 = no limit)

    // Torque jog (interactive manual torque, dead-man)
    stsTorqueJogActive  : BOOL;   // torque-jog engaged (held, or ramping back to 0 after release)
    stsTorqueJogMaxVel  : LREAL;  // [unit/s] active (retained) torque-jog overspeed trip; 0 = no trip

    // Position jog ("go to position") - discrete absolute move at the jog velocity/accel
    stsJogGotoBusy      : BOOL;   // TRUE while the go-to move is executing
    stsJogGotoDone      : BOOL;   // go-to move reached its target
    stsJogGotoPos       : LREAL;  // [unit] active/last go-to target position

    // Safety
    stsSTO              : BOOL;   // TRUE = STO not active (normal run), FALSE = STO active (drive torque cut imminent)
    stsSafetyInhibited  : BOOL;   // TRUE = motion inhibited by safety (STO active). Soft inhibit, NOT a fault:
                                  // blocks enable/motion, self-clears when STO restored (no reset needed)

    // Units / kinematics (NC carries no unit metadata - configured on fb_Axis)
    stsAxisType         : E_Axis_UnitType;  // eLinear / eRotary
    stsUnit             : STRING;           // position unit label (e.g. 'mm','deg'); velocity = unit + '/s'
    stsIsModulo         : BOOL;             // TRUE = axis is modulo: show stsModuloActPos, else stsActualPosition

    // Coordination
    stsExternalControl  : BOOL;   // axis yielded to external coordinator

    // Move list - mirrored from fb_Axis internal persistent moves for HMI display
    moves               : ARRAY[1..20] OF ST_Axis_MoveDefinition;
    // Live interlock status per move - shows which moves are currently executable
    moveInterlocks      : ARRAY[1..20] OF ST_Interlock_HMI_Interface;
END_STRUCT
END_TYPE

// ---- DUTs/fb_Axis/ST_Axis_MoveDefinition.TcDUT
// Move command struct. fb_Axis maintains a parallel ARRAY[1..20] OF fb_Interlock
// fed from each move's interlock field - giving each move its own live interlock FB.
TYPE ST_Axis_MoveDefinition :
STRUCT
    moveName     : STRING;             // display label - used in fault messages
    mode         : E_Axis_Mode;        // selects which MC block executes
    position     : LREAL;              // absolute position [unit] or relative distance [unit]
    velocity     : LREAL;              // [unit/s] - in eTorque mode: software max-velocity limit (0 = no limit)
    acceleration : LREAL;              // [unit/s²]
    deceleration : LREAL;              // [unit/s²]
    jerk         : LREAL;              // [unit/s³] - 0 = trapezoidal profile
    torque       : LREAL;              // [Nm or %] - used in eTorque mode
    torqueRamp   : LREAL;              // [torque unit/s] - used in eTorque mode, 0 = immediate
    cfgTorqueLimit : LREAL;            // [Nm or %] max |actual torque| allowed during this move (0 = no limit).
                                       //   Exceed → locked MC_Stop + fault 'Overtorque limit: <moveName>'.
                                       //   Applies to ALL modes (jam/collision protection); same units as ActTorque.
    direction    : MC_Direction;       // velocity/torque mode direction
    bufferMode   : E_Axis_BufferMode;  // Phase 1: only eAborting honored
    interlock    : ST_Interlock;       // move-level permissive - checked at execution
END_STRUCT
END_TYPE

// ---- DUTs/Camming/fb_CamCoupler/E_CamCoupler_State.TcDUT
// State of the couple/decouple sequence for one slave-master pair.
// Execution order of a couple: eIdle -> eYielding -> eSelecting -> eCoupling -> eCoupled.
// Execution order of a decouple: (engaged) -> eDecoupling -> eStopping -> eIdle (or eError on fault).
TYPE E_CamCoupler_State :
(
    eIdle       := 0,  // not coupled, waiting for a couple request
    eSelecting  := 1,  // MC_CamTableSelect running (register the verified table)
    eYielding   := 2,  // fb_Axis yielded; waiting for the slave to reach standstill before selecting
    eCoupling   := 3,  // MC_CamIn running (RampIn engage); waiting for InSync
    eCoupled    := 4,  // synchronized to the master via the cam (steady state)
    eDecoupling := 5,  // MC_CamOut running (disengage)
    eStopping   := 6,  // MC_Halt running to kill the retained slave velocity, then release the yield
    eError      := 7   // latched coupler error; requires cmdReset/inpReset
) INT;
END_TYPE

// ---- DUTs/Camming/fb_CamCoupler/ST_CamCoupler_HMI_Commands.TcDUT
// HMI -> PLC operator commands for the cam coupler.
// All ocmd* flags are self-clearing one-shots: the FB consumes and resets them the scan it sees them.
TYPE ST_CamCoupler_HMI_Commands :
STRUCT
    ocmdCouple          : BOOL;   // request engage (yield -> select -> cam-in)
    ocmdDecouple        : BOOL;   // request controlled decouple (cam-out -> stop -> release yield)
    ocmdReset           : BOOL;   // clear a latched coupler error and return to idle

    // Live cam-offset trim (no decouple): write the offset operand then pulse the matching set flag.
    ocmdSetMasterOffset : BOOL;   // apply ocmdMasterOffset as the new master offset (re-issues MC_CamIn)
    ocmdMasterOffset    : LREAL;  // [master unit] new cam master offset
    ocmdSetSlaveOffset  : BOOL;   // apply ocmdSlaveOffset as the new slave offset (re-issues MC_CamIn)
    ocmdSlaveOffset     : LREAL;  // [slave unit] new cam slave offset

    // Superimposed correction (no decouple): a bounded corrective move on top of the running cam.
    ocmdSuperImpose     : BOOL;   // run MC_MoveSuperImposed with the operands below
    ocmdSuperImposeDist : LREAL;  // [slave unit] corrective distance added on top of the cam
    ocmdSuperImposeVelo : LREAL;  // [slave unit/s] additional velocity for the correction
END_STRUCT
END_TYPE

// ---- DUTs/Camming/fb_CamCoupler/ST_CamCoupler_HMI_Config.TcDUT
// HMI-editable / commissioning mirror of the cam relationship.
// The live coupling values are wired to fb_CamCoupler VAR_INPUTs by the machine layer; this struct
// mirrors the configured defaults for commissioning display/editing (seeded from the cfg* defaults).
TYPE ST_CamCoupler_HMI_Config :
STRUCT
    masterOffset : LREAL;         // [master unit] default cam master offset
    slaveOffset  : LREAL;         // [slave unit]  default cam slave offset
    masterScale  : LREAL := 1.0;  // default master scaling
    slaveScale   : LREAL := 1.0;  // default slave scaling
    periodic     : BOOL;          // default MC_CamTableSelect periodicity
    tableId      : UDINT;         // default NC cam table id
END_STRUCT
END_TYPE

// ---- DUTs/Camming/fb_CamCoupler/ST_CamCoupler_HMI_Interface.TcDUT
// Public HMI interface for fb_CamCoupler - the struct an HMI binds.
// No HMIbaseDevice: fb_CamCoupler is standalone and does NOT extend abs_fb_Device.
TYPE ST_CamCoupler_HMI_Interface :
STRUCT
    Status   : ST_CamCoupler_HMI_Status;
    Commands : ST_CamCoupler_HMI_Commands;
    Config   : ST_CamCoupler_HMI_Config;
END_STRUCT
END_TYPE

// ---- DUTs/Camming/fb_CamCoupler/ST_CamCoupler_HMI_Status.TcDUT
// PLC -> HMI status for the cam coupler.
TYPE ST_CamCoupler_HMI_Status :
STRUCT
    stsState        : E_CamCoupler_State;  // current couple/decouple state
    stsCoupled      : BOOL;   // MC_CamIn.InSync - slave synchronized to the master via the cam
    stsBusy         : BOOL;   // a couple or decouple sequence is in progress
    stsError        : BOOL;   // latched coupler error (own error model - NOT an NC/axis fault)
    stsErrorText    : STRING;  // reason for the latched error

    stsVerified     : BOOL;   // echo of the incoming verified gate (from fb_CamTeach.stsVerified)
    stsTableId      : UDINT;  // NC cam table id in use for this coupling

    // Live cam relationship values (effective, latched at engage / updated by live trim)
    stsMasterOffset : LREAL;  // [master unit]
    stsSlaveOffset  : LREAL;  // [slave unit]
    stsMasterScale  : LREAL;  // master scaling
    stsSlaveScale   : LREAL;  // slave scaling
    stsPeriodic     : BOOL;   // MC_CamTableSelect periodicity in use
END_STRUCT
END_TYPE

// ---- DUTs/Camming/fb_CamTeach/E_CamTeach_Interp.TcDUT
// Interpolation strategy used by cmdConvert when building the motion function
// from the raw taught points. Stored raw, so this may change and be regenerated.
TYPE E_CamTeach_Interp :
(
    eLinear  := 0,   // straight segments between points (MOTIONFUNCTYPE_LINEAR)
    eCubicC1 := 1    // POLYNOM3 + central-difference slope -> C1-smooth cubic from position-only teaching
) INT;
END_TYPE

// ---- DUTs/Camming/fb_CamTeach/E_CamTeach_State.TcDUT
// Lifecycle state of one fb_CamTeach instance. Order/values are a CONTRACT:
// fb_CamTeach and any HMI depend on this exact ordering - do not reorder.
//   eIdle -cmdRecord-> eTeaching -cmdConvert-> eConverted -cmdDownload-> eDownloading -> eVerifying -> eVerified
//   save/load transition through eSaving/eLoading and return to the prior working state
//   any step error -> eError (stsErrorText); inpReset -> eIdle
TYPE E_CamTeach_State :
(
    eIdle        := 0,   // no operation in progress; working set may be empty or taught
    eTeaching    := 1,   // recording / editing raw points (working set is being built)
    eConverted   := 2,   // raw points post-processed and built into _mfPoints[], not yet downloaded
    eSaving      := 3,   // async file write in progress (fb_CamTeachFile)
    eLoading     := 4,   // async file read in progress (fb_CamTeachFile)
    eDownloading := 5,   // MC_WriteMotionFunction pushing _mfPoints[] to the NC table
    eVerifying   := 6,   // reading the table back and comparing to _mfPoints[]
    eVerified    := 7,   // table downloaded AND read-back-verified; stsVerified TRUE (gates coupling)
    eError       := 8    // last operation failed; see stsErrorText. inpReset returns to eIdle
) INT;
END_TYPE

// ---- DUTs/Camming/fb_CamTeach/ST_CamTeach_HMI_Commands.TcDUT
// HMI -> PLC operator commands for one cam-teach instance.
// Every ocmd* flag is a self-clearing one-shot: the HMI writes TRUE, fb_CamTeach
// acts on it and immediately writes it back to FALSE (same convention as fb_Axis).
// Operand fields (ocmd*Master / ocmd*Index / ...) are read on the scan the paired
// flag is seen, so the HMI must set them before (or with) the flag.
TYPE ST_CamTeach_HMI_Commands :
STRUCT
    // Record: append one raw taught point. The caller/HMI supplies BOTH values
    // (teach-by-value, not by axis) - master and slave are scalars.
    ocmdRecord          : BOOL;   // one-shot: append (ocmdRecordMaster, ocmdRecordSlave)
    ocmdRecordMaster    : LREAL;  // [master unit] master value for the recorded point
    ocmdRecordSlave     : LREAL;  // [slave unit]  slave value for the recorded point

    // Delete the most recently recorded point from the working set.
    ocmdDeleteLast      : BOOL;   // one-shot: remove last point

    // Spot-edit one existing point (offline, before convert/download).
    ocmdEditPoint       : BOOL;   // one-shot: overwrite point ocmdEditIndex
    ocmdEditIndex       : INT;    // 1..stsNumPoints target point index
    ocmdEditMaster      : LREAL;  // [master unit] new master value
    ocmdEditSlave       : LREAL;  // [slave unit]  new slave value

    // Empty the working set (returns toward eIdle).
    ocmdClear           : BOOL;   // one-shot: clear all taught points

    // Persist raw points -> file (async, via fb_CamTeachFile). ocmdFileName is the
    // bare file name; the directory is the FB's cfgFileDir concern.
    ocmdSave            : BOOL;   // one-shot: start async save
    ocmdFileName        : STRING; // file name to save to (also seeds/echoes Config.fileName)

    // File -> raw points (async). Loads from Config.fileName / last used name.
    ocmdLoad            : BOOL;   // one-shot: start async load

    // Post-process + build the motion function -> eConverted.
    ocmdConvert         : BOOL;   // one-shot: convert raw points to _mfPoints[]

    // Download _mfPoints[] to the NC table then read-back verify -> eVerified.
    ocmdDownload        : BOOL;   // one-shot: MC_WriteMotionFunction + verify

    // Online (live) point edit while cammed: update the slave of one point and apply
    // it at a defined master position (not immediately). Re-saves the file to stay truthful.
    ocmdEditOnline      : BOOL;   // one-shot: live edit point ocmdEditOnlineIndex
    ocmdEditOnlineIndex : INT;    // 1..stsNumPoints target point index
    ocmdEditOnlineSlave : LREAL;  // [slave unit] new slave value for the live edit

    // Clear a fault / return the FB to eIdle.
    ocmdReset           : BOOL;   // one-shot: reset (mirrors inpReset)
END_STRUCT
END_TYPE

// ---- DUTs/Camming/fb_CamTeach/ST_CamTeach_HMI_Config.TcDUT
// HMI-editable configuration for one cam-teach instance.
// These mirror the FB's cfg* settings so the operator can tune them from the screen;
// fb_CamTeach reads them when the paired command runs (e.g. fileName on save/load).
TYPE ST_CamTeach_HMI_Config :
STRUCT
    fileName    : STRING;              // bare file name to save to / load from (dir is the FB's concern)

    // ISO-8601 timestamp for the CSV header, supplied by the HMI. The wall clock is
    // not sampled in-scan, so the caller stamps 'created' (e.g. '2026-07-14T09:12:00').
    created     : STRING;              // 'created=' value written into the file metadata header

    // Editable tuning mirrors (applied on the relevant command / next convert):
    periodic    : BOOL;               // TRUE = periodic table (wrap velocity at the seam)
    interp      : E_CamTeach_Interp;  // interpolation strategy for cmdConvert
    smoothWindow: INT;                // moving-average window on master column (3-5; 0 = off)
    slaveName   : STRING;             // name of the slave this table teaches (goes into file header)
END_STRUCT
END_TYPE

// ---- DUTs/Camming/fb_CamTeach/ST_CamTeach_HMI_Interface.TcDUT
// Full HMI interface for one fb_CamTeach instance - the struct an HMI binds.
// Same nested Status / Commands / Config convention as ST_Axis_HMI_Interface, but with
// NO HMIbaseDevice: fb_CamTeach is a standalone library primitive and does NOT extend
// abs_fb_Device, so it carries its own error model (Status.stsError / stsErrorText).
TYPE ST_CamTeach_HMI_Interface :
STRUCT
    Status   : ST_CamTeach_HMI_Status;
    Commands : ST_CamTeach_HMI_Commands;
    Config   : ST_CamTeach_HMI_Config;
END_STRUCT
END_TYPE

// ---- DUTs/Camming/fb_CamTeach/ST_CamTeach_HMI_Status.TcDUT
// PLC -> HMI status for one cam-teach instance.
// sts* fields mirror the FB outputs plus curated readouts for the teach screen.
TYPE ST_CamTeach_HMI_Status :
STRUCT
    // Lifecycle
    stsState        : E_CamTeach_State;  // current state machine state (mirror of stsState output)
    stsNumPoints    : INT;               // number of raw points in the working set
    stsVerified     : BOOL;              // table downloaded AND read-back-verified (gates fb_CamCoupler)
    stsBusy         : BOOL;              // file / download / verify in progress

    // Error (own error model - this FB does not extend abs_fb_Device)
    stsError        : BOOL;              // an operation failed; latched until reset
    stsErrorText    : STRING;            // human-readable reason for stsError

    // File I/O readout (mirrors the fb_CamTeachFile sub-FB)
    stsFileBusy     : BOOL;              // async save/load in progress
    stsFileName     : STRING;            // file name of the last/active save or load

    // Last recorded pair - lets the HMI confirm what was just captured
    stsLastMaster   : LREAL;            // [master unit] master of the most recent recorded point
    stsLastSlave    : LREAL;            // [slave unit]  slave of the most recent recorded point

    // Config echo - what the FB is actually configured with (read-back of cfg*/Config)
    stsSlaveName    : STRING;            // name of the slave this table teaches
    stsPeriodic     : BOOL;              // TRUE = periodic table (velocity wraps at the seam)
    stsInterp       : E_CamTeach_Interp; // active interpolation strategy
    stsSmoothWindow : INT;               // moving-average window on master column (0 = off)
    stsTableId      : UDINT;             // NC motion-function table id bound to this instance

    // Bounded points preview - a tail of the working set for HMI spot-checking.
    // Intentionally NOT the full MAX_CAM_POINTS array: a 4096-deep LREAL array per
    // instance is too heavy to symbol-link to the HMI, so only the last few points
    // are exposed. stsPreviewCount says how many entries are valid (1..32).
    stsPreviewCount : INT;                          // number of valid entries in stsPreview (0..32)
    stsPreview      : ARRAY[1..32] OF ST_CamTeach_Point;  // tail (most recent) of the working set
END_STRUCT
END_TYPE

// ---- DUTs/Camming/fb_CamTeach/ST_CamTeach_Point.TcDUT
// One raw taught master->slave pair for THIS slave table.
// The file (CSV) stores these raw values; NC motion-function structs are
// regenerated from them on convert, so the interpolation strategy can change.
TYPE ST_CamTeach_Point :
STRUCT
    rMaster : LREAL;   // [master unit] strictly increasing after post-process (offset-zeroed, monotonic)
    rSlave  : LREAL;   // [slave unit]  taught slave position at rMaster
END_STRUCT
END_TYPE

// ---- DUTs/Devices/fb_Dev_StripLight_BannerWLS15Pro/E_BannerWLS15Pro_Animation.TcDUT
{attribute 'qualified_only'}
{attribute 'strict'}
{attribute 'to_string'}
// Run Mode animation, subindex 1 (219132 Rev. A, section 1.3.2).
TYPE E_BannerWLS15Pro_Animation :
(
    eOff             := 0,
    eSteady          := 1,
    eFlash           := 2,
    eTwoColorFlash   := 3,
    eTwoColorShift   := 4,
    eEndsSteady      := 5,
    eEndsFlash       := 6,
    eScroll          := 7,
    eCenterScroll    := 8,
    eBounce          := 9,
    eCenterBounce    := 10,
    eIntensitySweep  := 11,
    eTwoColorSweep   := 12,
    eSpectrum        := 13,
    eSingleEndSteady := 14,
    eSingleEndFlash  := 15
) BYTE;
END_TYPE

// ---- DUTs/Devices/fb_Dev_StripLight_BannerWLS15Pro/E_BannerWLS15Pro_Color.TcDUT
{attribute 'qualified_only'}
{attribute 'strict'}
{attribute 'to_string'}
// Run Mode Color 1 / Color 2, subindices 2 and 6 (219132 Rev. A, section 1.3.2).
// eCustom1 / eCustom2 render whatever was written to the device's custom
// colour parameters; the rest are fixed in firmware.
TYPE E_BannerWLS15Pro_Color :
(
    eGreen                  := 0,
    eRed                    := 1,
    eOrange                 := 2,
    eAmber                  := 3,
    eYellow                 := 4,
    eLimeGreen              := 5,
    eSpringGreen            := 6,
    eCyan                   := 7,
    eSkyBlue                := 8,
    eBlue                   := 9,
    eViolet                 := 10,
    eMagenta                := 11,
    eRose                   := 12,
    eDaylightWhite5000K     := 13,
    eCustom1                := 14,
    eCustom2                := 15,
    eIncandescentWhite2700K := 16,
    eWarmWhite3000K         := 17,
    eFluorescentWhite4100K  := 18,
    eNeutralWhite5700K      := 19,
    eCoolWhite6500K         := 20
) BYTE;
END_TYPE

// ---- DUTs/Devices/fb_Dev_StripLight_BannerWLS15Pro/E_BannerWLS15Pro_Direction.TcDUT
{attribute 'qualified_only'}
{attribute 'strict'}
{attribute 'to_string'}
// Run Mode direction / single-end animation location, subindex 10
// (219132 Rev. A, section 1.3.2).
TYPE E_BannerWLS15Pro_Direction :
(
    eUp   := 0,
    eDown := 1
) BYTE;
END_TYPE

// ---- DUTs/Devices/fb_Dev_StripLight_BannerWLS15Pro/E_BannerWLS15Pro_Intensity.TcDUT
{attribute 'qualified_only'}
{attribute 'strict'}
{attribute 'to_string'}
// Run Mode Color 1 / Color 2 Intensity, subindices 3 and 7 (219132 Rev. A,
// section 1.3.2). eCustom uses the device's custom intensity parameter.
TYPE E_BannerWLS15Pro_Intensity :
(
    eHigh   := 0,
    eLow    := 1,
    eMedium := 2,
    eOff    := 3,
    eCustom := 4
) BYTE;
END_TYPE

// ---- DUTs/Devices/fb_Dev_StripLight_BannerWLS15Pro/E_BannerWLS15Pro_PulsePattern.TcDUT
{attribute 'qualified_only'}
{attribute 'strict'}
{attribute 'to_string'}
// Run Mode pulse pattern, subindex 5 (219132 Rev. A, section 1.3.2).
// Only read by the flashing animations.
TYPE E_BannerWLS15Pro_PulsePattern :
(
    eNormal     := 0,
    eStrobe     := 1,
    eThreePulse := 2,
    eSOS        := 3,
    eRandom     := 4
) BYTE;
END_TYPE

// ---- DUTs/Devices/fb_Dev_StripLight_BannerWLS15Pro/E_BannerWLS15Pro_ScrollBounceStyle.TcDUT
{attribute 'qualified_only'}
{attribute 'strict'}
{attribute 'to_string'}
// Run Mode scroll/bounce style, subindex 8 (219132 Rev. A, section 1.3.2).
// Only read by the Scroll and Bounce animations.
TYPE E_BannerWLS15Pro_ScrollBounceStyle :
(
    eSolid  := 0,
    eTail   := 1,
    eRipple := 2
) BYTE;
END_TYPE

// ---- DUTs/Devices/fb_Dev_StripLight_BannerWLS15Pro/E_BannerWLS15Pro_Speed.TcDUT
{attribute 'qualified_only'}
{attribute 'strict'}
{attribute 'to_string'}
// Run Mode animation speed, subindex 4 (219132 Rev. A, section 1.3.2).
// eCustomFlashRate uses the device's custom flash rate parameter.
TYPE E_BannerWLS15Pro_Speed :
(
    eMedium          := 0,
    eFast            := 1,
    eSlow            := 2,
    eCustomFlashRate := 3
) BYTE;
END_TYPE

// ---- DUTs/Devices/fb_Dev_StripLight_BannerWLS15Pro/ST_Banner_WLS15PXRGB0220DSKQP_RunMode_Outputs.TcDUT
TYPE ST_Banner_WLS15PXRGB0220DSKQP_RunMode_Outputs :
STRUCT
	Direction 					: BYTE;
	Percent_Width_Of_Color_1 	: BYTE;
	Scroll_Bounce_Style			: BYTE;
	Color_2_Intensity			: BYTE;
	Color_2						: BYTE;
	Pulse_Pattern				: BYTE;
	Speed						: BYTE;
	Color_1_Intensity			: BYTE;
	Color_1						: BYTE;
	Animnation					: BYTE;
END_STRUCT
END_TYPE

// ---- DUTs/Devices/fb_Dev_XPendant/ST_XPendant_Axis.TcDUT
// One analog control broken into a DIRECTION trigger + a SPEED throttle, so it wires
// straight to a jog: Pos/Neg pick the jog direction, Throttle is the 0..100 % speed
// override. fb_Dev_XPendant derives one of these per stick axis and per trigger.
//   Sticks (bidirectional): Pos = up/right, Neg = down/left.
//   Triggers (one-sided):   Pos = pulled,   Neg always FALSE.
TYPE ST_XPendant_Axis :
STRUCT
    Value    : LREAL;   // raw gated deflection: sticks -1..1 (neg = down/left), triggers 0..1
    Pos      : BOOL;    // deflected + past cfgActivateThreshold (stick up/right; trigger pulled)
    Neg      : BOOL;    // deflected - past cfgActivateThreshold (stick down/left); FALSE for triggers
    Throttle : LREAL;   // 0..100 % speed = magnitude of deflection; 0 whenever neither Pos nor Neg
END_STRUCT
END_TYPE

// ---- DUTs/Devices/fb_Dev_XPendant/ST_XPendant_HMI_Interface.TcDUT
// HMI interface for fb_Dev_XPendant (bound as <instance>.HMI).
// No Commands/Config sub-structs: the pendant is an input-only device — its
// enable/disable lives in the IPC service (surface C), and config (feed timeout)
// is instantiation-time via FB_Init/cfgFeedTimeout, not operator-editable.
TYPE ST_XPendant_HMI_Interface :
STRUCT
    // Inherited base-device HMI values (deviceName, enabled, stsInAuto, stsFaulted,
    // stsFaultDescription, interlock). Populated from abs_fb_Device.
    HMIbaseDevice : ST_Device_HMI_Interface;
    Status        : ST_XPendant_HMI_Status;
END_STRUCT
END_TYPE

// ---- DUTs/Devices/fb_Dev_XPendant/ST_XPendant_HMI_Status.TcDUT
// Read-only pendant status for the HMI. Mirrors fb_Dev_XPendant's GATED sts*
// outputs (all idle unless stsConnected) plus the liveness diagnostics.
TYPE ST_XPendant_HMI_Status :
STRUCT
    stsConnected : BOOL;    // controller present AND feed alive AND enabled
    stsFeedAlive : BOOL;    // service watchdog fresh (diagnostic: FALSE + Connected claimed = service died)
    stsActive    : BOOL;    // inpActive AND stsConnected — pendant in service and usable now
    stsInService : BOOL;    // mirror of inpActive (supervision: pendant expected) — read by the IPC service

    stsBtnA      : BOOL;
    stsBtnB      : BOOL;
    stsBtnX      : BOOL;
    stsBtnY      : BOOL;
    stsBumpL     : BOOL;
    stsBumpR     : BOOL;
    stsStart     : BOOL;
    stsBack      : BOOL;
    stsThumbL    : BOOL;
    stsThumbR    : BOOL;

    stsDpadUp    : BOOL;
    stsDpadDown  : BOOL;
    stsDpadLeft  : BOOL;
    stsDpadRight : BOOL;

    // Analogs as direction + speed pairs (mirror of the FB outputs).
    stsLeftStickX  : ST_XPendant_Axis;
    stsLeftStickY  : ST_XPendant_Axis;
    stsRightStickX : ST_XPendant_Axis;
    stsRightStickY : ST_XPendant_Axis;
    stsTriggerL    : ST_XPendant_Axis;
    stsTriggerR    : ST_XPendant_Axis;
END_STRUCT
END_TYPE

// ---- DUTs/Devices/fb_Dev_XPendant/ST_XPendant_In.TcDUT
// Written over ADS by the lhmi `xpendant` sidecar app (lhmi-core apps/xpendant),
// which reads a USB Xbox controller on the IPC. This is a RAW EXTERNAL MIRROR, so
// members are unprefixed PascalCase (CONVENTIONS.md §2 exception) — the member
// names ARE the ADS write contract: the service writes <instance>.inpPad.<member>.
// PLC logic must never write into this struct.
TYPE ST_XPendant_In :
STRUCT
    Connected : BOOL;   // controller present AND service feeding
    Watchdog  : UINT;   // rolls 0..65535 every ~500 ms — stale => treat as disconnected

    // Face / shoulder / menu buttons
    BtnA      : BOOL;
    BtnB      : BOOL;
    BtnX      : BOOL;
    BtnY      : BOOL;
    BumpL     : BOOL;   // left bumper (LB)
    BumpR     : BOOL;   // right bumper (RB)
    Start     : BOOL;
    Back      : BOOL;
    ThumbL    : BOOL;   // left-stick click (L3)
    ThumbR    : BOOL;   // right-stick click (R3)

    // D-pad
    DpadUp    : BOOL;
    DpadDown  : BOOL;
    DpadLeft  : BOOL;
    DpadRight : BOOL;

    // Analog sticks: -1.0 .. 1.0, dead zone applied by the service, up/right = +
    StickLX   : LREAL;
    StickLY   : LREAL;
    StickRX   : LREAL;
    StickRY   : LREAL;

    // Analog triggers: 0.0 .. 1.0
    TrigL     : LREAL;
    TrigR     : LREAL;
END_STRUCT
END_TYPE

// ---- DUTs/Common/ST_Bits.TcDUT
TYPE ST_Bits :
STRUCT
	Bit1:BIT;
	Bit2:BIT;
	Bit3:BIT;
	Bit4:BIT;
	Bit5:BIT;
	Bit6:BIT;
	Bit7:BIT;
	Bit8:BIT;
	Bit9:BIT;
	Bit10:BIT;
	Bit11:BIT;
	Bit12:BIT;
	Bit13:BIT;
	Bit14:BIT;
	Bit15:BIT;
	Bit16:BIT;
END_STRUCT
END_TYPE

// ---- DUTs/Devices/fb_Dev_ControlValve_Modulating/ST_ControlValve_Modulating_HMI_Interface.TcDUT
TYPE ST_ControlValve_Modulating_HMI_Interface :
STRUCT
	HMIbaseDevice		: ST_Device_HMI_Interface;
	stsValveFeedback	: LREAL;	// position feedback from device
	ocmdValvePosition	: LREAL;    // operator command - valve position
	stsValvePosition	: LREAL;    // actual command - valve position
END_STRUCT
END_TYPE

// ---- DUTs/fb_IO_EL6751_Bus_Status/ST_EL6751_Bus_State.TcDUT
TYPE ST_EL6751_Bus_State :
STRUCT
	GlobalState0	:	UINT;
	GlobalState2	:	U_UINT16;
	GlobalState3	:	UINT;
END_STRUCT
END_TYPE

// ---- DUTs/fb_IO_EL6751_Bus_Status/ST_EL6751_Bus_State_Parsed.TcDUT
TYPE ST_EL6751_Bus_State_Parsed :
STRUCT
	stsCANDeviceState				:STRING;
	stsCANControllerBusOff			:BOOL;
	stsCANControllerWarningLimit	:BOOL;
	stsRxQueueOverrun				:BOOL;
	stsCANSendError					:BOOL;
	stsCANQueueIntRxOverflow		:BOOL;
	stsCANQueueIntTxOverflow		:BOOL;
	stsSyncToggle					:BOOL;
	stsBusLoad						:UINT;
END_STRUCT
END_TYPE

// ---- DUTs/fb_Interlock/ST_Interlock.TcDUT
TYPE ST_Interlock :
STRUCT
	conditions	: ARRAY[1..10] OF BOOL := [1,1,1,1,1,1,1,1,1,1];
	descriptions	: ARRAY[1..10] OF STRING := ['N/A','N/A','N/A','N/A','N/A','N/A','N/A','N/A','N/A','N/A'];
END_STRUCT
END_TYPE

// ---- DUTs/fb_Permissive/ST_Permissive.TcDUT
// Configuration for fb_Permissive: the conditions that must ALL be true, plus the operator-
// facing text for each. Mirrors ST_Interlock deliberately — same shape, same bound, same defaults,
// spelled the same literal way — so the two are interchangeable to read and a set of conditions can
// move between them.
//
// TEN SLOTS, HARDCODED. The bound is a literal here and in every FOR loop that walks it, per
// CONVENTIONS §5: a library DUT cannot reference a GVL for its sizing, because a DUT is a type and
// has no interface to receive one through. Raising the capacity means editing this bound and
// fb_Permissive's loops together — visible in review, which a GVL edit three files away is not.
//
// conditions DEFAULT TO TRUE. That is the load-bearing default: a permissive with only three
// of its ten slots wired must be satisfied by those three, not blocked forever by seven unwired
// FALSEs. Wire what applies and leave the rest.
//
// descriptions default to 'N/A' so an unwired slot never renders as blank on the HMI. Write real
// text for every slot you DO wire — that text is the operator's answer to "why won't it start",
// and an unnamed unmet condition is a dead end for them.
TYPE ST_Permissive :
STRUCT
    conditions      : ARRAY[1..10] OF BOOL := [1,1,1,1,1,1,1,1,1,1];
    descriptions    : ARRAY[1..10] OF STRING := ['N/A','N/A','N/A','N/A','N/A','N/A','N/A','N/A','N/A','N/A'];
END_STRUCT
END_TYPE

// ---- DUTs/fb_Permissive/ST_Permissive_HMI_Interface.TcDUT
// HMI face of fb_Permissive. Bind <instance>.HMI.* — the shared lhmi `PermissiveList` component
// renders exactly this struct, so any permissive anywhere (a device's start conditions, a
// MachineFlow transition gate, a machine-level ready check) gets the same operator view for free.
//
// There is deliberately NO first-out field here. First-out answers "which condition dropped and
// caused the trip", which only means something for an interlock: it faults instantly, so the
// condition that went first is the cause and the later ones are consequences. A permissive never
// trips - it is evaluated at the moment something asks to proceed, and every unmet condition is
// equally and simultaneously the reason. So this struct carries the SET (stsConditions) plus a
// count, and the HMI shows all of them rather than nominating a misleading headline.
//
// There is deliberately NO BYPASS field either. A permissive is not a safety function, so the
// temptation is to say a bypass is harmless here — but it is the one control that can make an
// unsatisfied gate report itself satisfied, and a sequence that advances on a forced permissive
// fails somewhere downstream where nothing explains why. Hold the conditions or do not; there is
// no third answer to publish. (fb_Interlock's inpGlobalBypass is a different case: an interlock
// stops a running machine, so commissioning needs a documented way to move it.)
//
// Bounds are literals, per CONVENTIONS §5 — matched to ST_Permissive's ten slots. Plain STRING is
// STRING(80), the same width the descriptions carry there.
TYPE ST_Permissive_HMI_Interface :
STRUCT
    stsPermissiveOK     : BOOL;     // TRUE when every condition is met
    stsConditions       : ARRAY[1..10] OF BOOL;
    stsDescriptions     : ARRAY[1..10] OF STRING;
    stsUnmetCount       : INT;      // how many are unmet — 0 when satisfied
    stsPermissiveName   : STRING;   // set via the cfgName property
END_STRUCT
END_TYPE

// ---- DUTs/fb_Interlock/ST_Interlock_HMI_Interface.TcDUT
TYPE ST_Interlock_HMI_Interface :
STRUCT
	stsInterlockOK				: BOOL;
	stsConditions				: ARRAY[1..10] OF BOOL;
	stsInterlockDescriptions 	: ARRAY[1..10] OF STRING;
	stsInterlockName			: STRING;

END_STRUCT
END_TYPE

// ---- DUTs/fb_Machine/ST_Machine_HMI_Interface.TcDUT
TYPE ST_Machine_HMI_Interface :
STRUCT
	inpReset				: BOOL;
	inpStop					: BOOL;
	inpStart				: BOOL;
	inpAuto					: BOOL;
	inpManual				: BOOL;
	inpInterlockBypass		: BOOL;
	inpAbort				: BOOL;
	inpPause				: BOOL;
	inpClearMachineLog		: BOOL;
	stsStopped				: BOOL;
	stsStarted				: BOOL;
	stsStartEnable			: BOOL;
	stsStartReady			: BOOL;
	stsInAuto				: BOOL;
	stsAutoEnable			: BOOL;
	stsInManual				: BOOL;
	stsInterlockBypassed	: BOOL;
	stsPaused				: BOOL;
	stsPausing				: BOOL;
	stsPauseEnable			: BOOL;
	stsInterlocksBypassed	: BOOL;
	stsMachineName			: T_MaxString;
	stsHeartBeat			: BOOL;			// toggles 500ms on / 500ms off - HMI frozen-data watchdog (binds machine.heartbeat)
END_STRUCT
END_TYPE

// ---- DUTs/Comm/ST_Modbus_Commands.TcDUT
TYPE ST_Modbus_Commands :
STRUCT
	ReadRegisters			: FB_MBReadRegs;
	ReadInputs				: FB_MBReadInputs;
	WriteSingleCoil			: FB_MBWriteSingleCoil;
	WriteSingleRegister		: FB_MBWriteSingleReg;
	WriteRegisters			: FB_MBWriteRegs;
END_STRUCT
END_TYPE

// ---- DUTs/Comm/ST_Modbus_Device_Config.TcDUT
TYPE ST_Modbus_Device_Config :
STRUCT
	cfgIP_address	: STRING(15);
	cfgTCPPort		: UINT;
	cfgUnitID		: BYTE;
	cfgTimeout		: TIME;
END_STRUCT
END_TYPE

// ---- DUTs/Common/U_ByteToLReal.TcDUT
TYPE U_ByteToLReal :
UNION
	bytes : ARRAY [1..4] OF  BYTE;
	value	:REAL;
END_UNION
END_TYPE

// ---- DUTs/Common/U_UINT16.TcDUT
TYPE U_UINT16 :
UNION
	Bits : ARRAY [1..1] OF  ST_Bits;
	Num : UINT;
END_UNION
END_TYPE

// ---- DUTs/Common/U_USINT.TcDUT
TYPE U_USINT :
UNION
	Bits : ARRAY [1..1] OF  ST_Bits;
	Num : USINT;
END_UNION
END_TYPE

// ---- GVLs/GVL_Cam.TcGVL
// Shared constants for the cam-teach subsystem (fb_CamTeach / fb_CamTeachFile).
// Kept in a GVL so the working-point array bound is a single source of truth
// across the FB, its persistence sub-FB, and any pre-created NC tables.
VAR_GLOBAL CONSTANT
    MAX_CAM_POINTS : INT := 4096;   // >= 360/rev x 7 revs + margin; array bound for cam point buffers
END_VAR

// ---- Version/Global_Version.TcGVL
{attribute 'TcGenerated'}
{attribute 'no-analysis'}
{attribute 'linkalways'}
// This function has been automatically generated from the project information.
VAR_GLOBAL CONSTANT
	{attribute 'const_non_replaced'}
	stLibVersion_LPLC : ST_LibVersion := (iMajor := 2, iMinor := 2, iBuild := 0, iRevision := 0, nFlags := 0, sVersion := '2.2.0');
END_VAR

// ---- POUs/FBs/Camming/fb_CamTeach.TcPOU
// fb_CamTeach - reusable, machine-agnostic teach/manage engine for ONE NC cam table
// (the master->slave relationship of a single slave). It records raw taught points,
// persists them to file (source of truth), post-processes + converts them into an NC
// motion function, downloads that function to a pre-created NC table and read-back
// verifies it, and exposes a per-table 'verified' flag that gates downstream coupling
// (fb_CamCoupler). It NEVER issues axis motion - its job ends at a verified table.
//
// Standalone library primitive: does NOT extend abs_fb_Device. It carries its OWN error
// model (stsError / stsErrorText, via the private setError) - never setFault, which does
// not exist here. Teach-by-value: cmdRecord takes scalar master/slave, not an AXIS_REF,
// so the caller decides where the values come from (real axis, virtual master, accumulator).
//
// Async work (file I/O, download, verify, online edit) is multi-scan. File I/O is isolated
// in the sub-FB fb_CamTeachFile, driven every scan with the working point array. Convert is
// SYNCHRONOUS (a pure, bounded compute). Download/verify + online edit are ASYNCHRONOUS
// state machines driven cyclically in the body.
//
// Convert is intentionally in-place: post-processing zeroes/compacts/smooths the working set
// (the design doc's "compact the array"), so raw points should be SAVED BEFORE convert (or
// reloaded) if the untouched raw values are needed - the file is the raw source of truth.
//
// NOTE: cfgMasterUnit is NOT in the design doc's cfg list; it is added here because the CSV
// header carries a machine-specific master unit that fb_CamTeachFile.cmdSave requires. See report.
FUNCTION_BLOCK fb_CamTeach
VAR_INPUT
    inpReset : BOOL;                 // level: while TRUE, hold the FB reset to E_CamTeach_State.eIdle (mirrors cmdReset)
END_VAR

VAR_OUTPUT
    stsState     : E_CamTeach_State;  // lifecycle state (mirror of _state)
    stsNumPoints : INT;               // number of raw points in the working set
    stsVerified  : BOOL;              // table downloaded AND read-back-verified - gates fb_CamCoupler
    stsBusy      : BOOL;              // file / download / verify / online edit in progress
    stsError     : BOOL;              // an operation failed; latched until reset
    stsErrorText : STRING;            // human-readable reason for stsError
END_VAR

VAR
    // Public HMI interface - the struct an HMI (e.g. lhmi) binds
    HMI      : ST_CamTeach_HMI_Interface;

    // Raw taught points (working set) + count and lifecycle state
    _points  : ARRAY[1..MAX_CAM_POINTS] OF ST_CamTeach_Point;
    _n       : INT;
    _state   : E_CamTeach_State;

    // NC motion-function table this instance owns (pre-created under Motion -> Tables).
    _tableId   : UDINT;               // NC cam-table id, set via cfgTableId / FB_Init (0 = unbound)
    // VERIFY against installed Tc2_MC2_Camming / TF5050: the struct name MC_MotionFunctionPoint
    // and ALL of its field names/types are library-version dependent (see cmdConvert).
    _mfPoints  : ARRAY[1..MAX_CAM_POINTS] OF MC_MotionFunctionPoint;   // VERIFY (struct name)
    _mcSelect  : Tc2_MC2_Camming.MC_CamTableSelect; // download: CREATES the NC table and fills it from _mfPoints
    _mcRead    : MC_ReadMotionFunctionPoint;     // VERIFY (block name + I/O) - per-point read-back
    _mcWritePt : MC_WriteMotionFunctionPoint;    // VERIFY (block name + I/O) - online single-point edit
    _mcOnline  : MC_SetCamOnlineChangeMode;      // VERIFY (block name + I/O + mode enum) - online change timing
    _readPt    : MC_MotionFunctionPoint;         // read-back target for MC_ReadMotionFunctionPoint (VAR_IN_OUT Point)
    _camWriteRef : MC_CAM_REF;                   // table descriptor for MC_CamTableSelect (pArray -> _mfPoints)

    _file : fb_CamTeachFile;          // isolated async CSV persistence sub-FB

    // Configuration backing (FB_Init + cfg* properties, per the fb_Axis pattern)
    _slaveName    : STRING;
    _periodic     : BOOL;
    _interp       : E_CamTeach_Interp;
    _smoothWindow : INT;                              // moving-average window on master column (0 = off)
    _fileDir      : STRING := 'C:\_MachineConfig\CamTables';
    _masterUnit   : STRING := 'mm';                  // CSV header master unit (added cfg - see header note)

    // Download / verify async sub-steps
    _dlStep    : INT;                                // sub-step inside eVerifying (0 = reading, 1 = advance)
    _verifyIdx : INT := 1;                           // point index being read back / compared
    _verifyEps : LREAL := 0.001;                     // read-back comparison tolerance (absolute)

    // Online-edit async sequence
    _onlineStep     : INT;                           // 0 idle; 10 set change-mode; 20 write pt; 30 advance
    _onlineIdx      : INT := 1;                       // point being edited online
    _onlineWriteIdx : INT := 1;                       // cursor over affected points (idx-1 .. idx+1)
    _onlineHi       : INT := 1;                       // last affected point index (min(_n, idx+1))
    _onlineSaveReq  : BOOL;                           // re-save the file after the online write completes

    // HMI readouts
    _lastMaster : LREAL;                             // master of the most recent recorded point
    _lastSlave  : LREAL;                             // slave  of the most recent recorded point
    _fileName   : STRING;                            // file name of the last save/load

    _returnState  : E_CamTeach_State;                // resting state to return to after eSaving
    _hmiCfgLoaded : BOOL;                            // HMI.Config seeded from cfg once

    _previewCount : INT;                             // valid entries in HMI.Status.stsPreview (0..32)
    _i            : INT;                             // loop index (body only)
END_VAR

// ── 1. Drive the persistence sub-FB every scan ───────────────────────────────
// It reads/writes the shared working buffer via VAR_IN_OUT; cmd* on _file only ARM ops.
_file(points := _points);

// ── 2. Reset handling ────────────────────────────────────────────────────────
// inpReset is level-driven: hold reset while TRUE (idempotent - clears error, returns to idle).
IF inpReset THEN
    cmdReset();
END_IF

// ── 3. HMI commands ──────────────────────────────────────────────────────────
// Seed the HMI.Config mirror once from the configured defaults; thereafter operator edits
// to the tuning mirrors flow back into the cfg backing so the next convert/save uses them
// (same seed-once-then-track convention as fb_Axis). 'created' is read live in cmdSave.
IF NOT _hmiCfgLoaded THEN
    HMI.Config.slaveName    := _slaveName;
    HMI.Config.periodic     := _periodic;
    HMI.Config.interp       := _interp;
    HMI.Config.smoothWindow := _smoothWindow;
    HMI.Config.fileName     := _fileName;
    _hmiCfgLoaded := TRUE;
ELSE
    _slaveName := HMI.Config.slaveName;
    _periodic  := HMI.Config.periodic;
    _interp    := HMI.Config.interp;
    IF HMI.Config.smoothWindow >= 0 THEN
        _smoothWindow := HMI.Config.smoothWindow;
    END_IF
END_IF

// Self-clearing one-shot command dispatch (same convention as fb_Axis section 3):
// on seeing an ocmd* flag, immediately write it back FALSE, then call the matching method.
IF HMI.Commands.ocmdReset THEN
    HMI.Commands.ocmdReset := FALSE;
    cmdReset();
END_IF

IF HMI.Commands.ocmdRecord THEN
    HMI.Commands.ocmdRecord := FALSE;
    cmdRecord(HMI.Commands.ocmdRecordMaster, HMI.Commands.ocmdRecordSlave);
END_IF

IF HMI.Commands.ocmdDeleteLast THEN
    HMI.Commands.ocmdDeleteLast := FALSE;
    cmdDeleteLast();
END_IF

IF HMI.Commands.ocmdEditPoint THEN
    HMI.Commands.ocmdEditPoint := FALSE;
    cmdEditPoint(HMI.Commands.ocmdEditIndex, HMI.Commands.ocmdEditMaster, HMI.Commands.ocmdEditSlave);
END_IF

IF HMI.Commands.ocmdClear THEN
    HMI.Commands.ocmdClear := FALSE;
    cmdClear();
END_IF

IF HMI.Commands.ocmdSave THEN
    HMI.Commands.ocmdSave := FALSE;
    HMI.Config.fileName := HMI.Commands.ocmdFileName;   // ocmdFileName seeds/echoes Config.fileName
    cmdSave(HMI.Commands.ocmdFileName);
END_IF

IF HMI.Commands.ocmdLoad THEN
    HMI.Commands.ocmdLoad := FALSE;
    cmdLoad(HMI.Commands.ocmdFileName);
END_IF

IF HMI.Commands.ocmdConvert THEN
    HMI.Commands.ocmdConvert := FALSE;
    cmdConvert();
END_IF

IF HMI.Commands.ocmdDownload THEN
    HMI.Commands.ocmdDownload := FALSE;
    cmdDownload();
END_IF

IF HMI.Commands.ocmdEditOnline THEN
    HMI.Commands.ocmdEditOnline := FALSE;
    cmdEditOnline(HMI.Commands.ocmdEditOnlineIndex, HMI.Commands.ocmdEditOnlineSlave);
END_IF

// ── 4. Async state machine progression ───────────────────────────────────────
// Reacts to the results (from LAST scan's block calls) of the file sub-FB and the MC blocks,
// then section 4c drives the blocks for THIS scan. Convert is synchronous (in cmdConvert).
CASE _state OF

    eSaving:
        IF _file.stsError THEN
            setError(CONCAT('File save failed: ', _file.stsErrorText));
        ELSIF _file.stsDone THEN
            _state := _returnState;                 // save leaves the data unchanged -> prior state
        END_IF

    eLoading:
        IF _file.stsError THEN
            setError(CONCAT('File load failed: ', _file.stsErrorText));
        ELSIF _file.stsDone THEN
            _n          := _file.stsNumPointsLoaded;
            stsVerified := FALSE;                    // loaded points need re-convert + re-download
            IF _n < 2 THEN
                setError('Loaded file has too few points (need >= 2)');
            ELSE
                _state := eTeaching;
            END_IF
        END_IF

    eDownloading:
        IF _mcSelect.Error THEN
            setError(CONCAT('Table create error: ', UDINT_TO_STRING(_mcSelect.ErrorID)));
        ELSIF _mcSelect.Done THEN
            _verifyIdx := 1;
            _dlStep    := 0;
            _state     := eVerifying;
        END_IF

    eVerifying:
        CASE _dlStep OF
            0:  // waiting for the read-back of point _verifyIdx (compare within _verifyEps)
                IF _mcRead.Error THEN
                    stsVerified := FALSE;
                    setError(CONCAT('Table read error: ', UDINT_TO_STRING(_mcRead.ErrorID)));
                ELSIF _mcRead.Done THEN
                    // Read-back point is delivered via the VAR_IN_OUT Point (-> _readPt), compared within _verifyEps.
                    IF   ABS(_readPt.MasterPos - _mfPoints[_verifyIdx].MasterPos) > _verifyEps
                      OR ABS(_readPt.SlavePos  - _mfPoints[_verifyIdx].SlavePos)  > _verifyEps THEN
                        stsVerified := FALSE;
                        setError(CONCAT('Verify mismatch at point ', INT_TO_STRING(_verifyIdx)));
                    ELSE
                        _dlStep := 1;               // point OK -> deassert one scan, then advance
                    END_IF
                END_IF
            1:  // deassert scan complete: step to the next point, or finish
                _verifyIdx := _verifyIdx + 1;
                IF _verifyIdx > _n THEN
                    stsVerified := TRUE;            // downloaded AND read-back-verified -> gates coupling
                    _state      := eVerified;
                ELSE
                    _dlStep := 0;
                END_IF
        END_CASE

END_CASE

// ── 4b. Online-edit write sequence (MC_SetCamOnlineChangeMode + MC_WriteMotionFunctionPoint) ─
// Runs independently of _state (a live edit while the table is in use); stsBusy reflects it.
CASE _onlineStep OF
    10:  // configure the online-change mode (apply at a defined master position, not immediately)
        IF _mcOnline.Error THEN
            setError(CONCAT('Online change-mode error: ', UDINT_TO_STRING(_mcOnline.ErrorID)));
        ELSIF _mcOnline.Done THEN
            _onlineStep := 20;
        END_IF
    20:  // writing affected point _onlineWriteIdx
        IF _mcWritePt.Error THEN
            setError(CONCAT('Online point write error: ', UDINT_TO_STRING(_mcWritePt.ErrorID)));
        ELSIF _mcWritePt.Done THEN
            _onlineStep := 30;                       // deassert one scan, then advance
        END_IF
    30:  // advance to the next affected point (idx-1 .. idx+1), or finish + re-save
        _onlineWriteIdx := _onlineWriteIdx + 1;
        IF _onlineWriteIdx > _onlineHi THEN
            _onlineStep     := 0;
            _onlineWriteIdx := 1;                    // keep the cursor in-bounds (4c reads _mfPoints[cursor])
            IF _onlineSaveReq AND _fileName <> '' THEN
                _onlineSaveReq := FALSE;
                cmdSave(_fileName);                  // keep the file truthful after a live edit
            END_IF
        ELSE
            _onlineStep := 20;
        END_IF
END_CASE

// ── 4c. Drive the Tc2_MC2_Camming blocks (called every scan; Execute gated by state) ─────
// Download: MC_CamTableSelect CREATES NC table _tableId and fills it with _mfPoints[1.._n] (TF5050
// manual 5.1: "creates a new table and simultaneously fills it with data provided by the PLC").
// NOT MC_WriteMotionFunction: that only rewrites points of a table already loaded in the NC - on a
// table that does not exist yet (or an empty System Manager table) the NC answers ADS 0x701
// "service not supported" (seen on a test rig, 2026-10-18). The table id must NOT also be a table defined in the
// System Manager. Periodicity is fixed here, at creation (MC_CamIn has no periodic input).
// MC_CAM_REF must FULLY describe the source buffer (an unset TableType -> 19249). Motion function =
// 1 column; NoOfRows = point count; ArraySize = the bytes of those points, so size, rows and columns
// agree.
_camWriteRef.pArray      := ADR(_mfPoints[1]);
_camWriteRef.ArraySize   := INT_TO_UDINT(_n) * SIZEOF(_mfPoints[1]);
_camWriteRef.TableType   := MC_TABLETYPE_MOTIONFUNCTION;
_camWriteRef.NoOfColumns := 1;
_camWriteRef.NoOfRows    := INT_TO_UDINT(_n);
_mcSelect(
    Execute    := (_state = eDownloading),
    Periodic   := _periodic,
    CamTableID := _tableId,
    CamTable   := _camWriteRef                                          // VAR_IN_OUT: fully-described MC_CAM_REF
);

// Verify: per-point read-back of point _verifyIdx (Execute pulses low between points).
// VERIFY: block name, CamTableID/PointIndex input names, and the MotionFunctionPoint output.
_mcRead(
    Execute    := (_state = eVerifying) AND (_dlStep = 0),
    CamTableID := _tableId,                                              // VERIFY: MC_CAM_ID type
    PointID    := INT_TO_UDINT(_verifyIdx),                             // point-index input (MC_MotionFunctionPoint_ID)
    Point      := _readPt                                                // VAR_IN_OUT: read-back point lands here
);

// Online single-point edit: write the changed/affected point live.
// VERIFY: block name + MotionFunctionPoint input struct name.
_mcWritePt(
    Execute    := (_onlineStep = 20),
    CamTableID := _tableId,                                              // VERIFY: MC_CAM_ID type
    PointID    := _mfPoints[_onlineWriteIdx].PointIndex,                // MC_MotionFunctionPoint_ID of the edited point
    Point      := _mfPoints[_onlineWriteIdx]                             // VAR_IN_OUT: point data to write
);

// Online change mode: apply the live edit at a DEFINED master position (not immediately),
// so editing the segment the slave is currently traversing does not step the setpoint.
// VERIFY: block name, mode enum name/value, and how the defined master position is specified -
// some versions apply "on next cam cycle" (the period seam) instead of an explicit MasterPos.
_mcOnline(
    Execute            := (_onlineStep = 10),
    CamTableID         := _tableId,                                     // VERIFY: MC_CAM_ID type
    ActivationMode     := MC_CAMACTIVATION_ATMASTERAXISPOS,             // apply at a defined master axis position
    ActivationPosition := 0.0                                           // table origin / seam
);

// ── 5. Outputs + HMI status ──────────────────────────────────────────────────
stsState     := _state;
stsNumPoints := _n;
stsBusy      := _file.stsBusy
                OR (_state = eSaving) OR (_state = eLoading)
                OR (_state = eDownloading) OR (_state = eVerifying)
                OR (_onlineStep <> 0);
// stsVerified / stsError / stsErrorText are maintained by the command + verify logic above.

// Bounded preview: the most-recent tail of the working set (<= 32 points) for HMI spot-checks.
_previewCount := _n;
IF _previewCount > 32 THEN
    _previewCount := 32;
END_IF
FOR _i := 1 TO 32 DO
    IF _i <= _previewCount THEN
        HMI.Status.stsPreview[_i] := _points[_n - _previewCount + _i];
    ELSE
        HMI.Status.stsPreview[_i].rMaster := 0.0;
        HMI.Status.stsPreview[_i].rSlave  := 0.0;
    END_IF
END_FOR

HMI.Status.stsState        := _state;
HMI.Status.stsNumPoints    := _n;
HMI.Status.stsVerified     := stsVerified;
HMI.Status.stsBusy         := stsBusy;
HMI.Status.stsError        := stsError;
HMI.Status.stsErrorText    := stsErrorText;
HMI.Status.stsFileBusy     := _file.stsBusy;
HMI.Status.stsFileName     := _fileName;
HMI.Status.stsLastMaster   := _lastMaster;
HMI.Status.stsLastSlave    := _lastSlave;
HMI.Status.stsSlaveName    := _slaveName;         // config echo (read-back of cfg*/Config)
HMI.Status.stsPeriodic     := _periodic;
HMI.Status.stsInterp       := _interp;
HMI.Status.stsSmoothWindow := _smoothWindow;
HMI.Status.stsTableId      := _tableId;
HMI.Status.stsPreviewCount := _previewCount;

// Append one raw taught point (caller supplies BOTH scalars - teach by value, not by axis).
// Bounds-checked against MAX_CAM_POINTS. Recording invalidates any verified table and moves
// to eTeaching. Rejected QUIETLY while an async op is running or while errored.
METHOD PUBLIC cmdRecord : BOOL
VAR_INPUT
    rMaster : LREAL;   // [master unit]
    rSlave  : LREAL;   // [slave unit]
END_VAR
cmdRecord := FALSE;
IF isBusy() OR stsError THEN
    RETURN;
END_IF

IF _n >= MAX_CAM_POINTS THEN
    setError('Record: cam point buffer full');
    RETURN;
END_IF

_n := _n + 1;
_points[_n].rMaster := rMaster;
_points[_n].rSlave  := rSlave;
_lastMaster := rMaster;
_lastSlave  := rSlave;
stsVerified := FALSE;                 // editing/recording clears verified
_state      := eTeaching;
cmdRecord   := TRUE;
END_METHOD

// Remove the most recently recorded point. Clears verified. Rejected QUIETLY while busy/errored.
METHOD PUBLIC cmdDeleteLast : BOOL
cmdDeleteLast := FALSE;
IF isBusy() OR stsError THEN
    RETURN;
END_IF

